FUNCTION_BLOCK "FB_GRAPH_PressDemoAuto"   // FB100, GRAPH
VERSION : 0.1
// stored: AcknowledgeErrorsRequired true, AutoNumber true, GraphVersion 6.0, InitialValuesAcquisition false, IsIECCheckEnabled false, LanguageInNetworks LAD, LockOperatingMode false, PermanentILProcessingInMANMode false, SetENOAutomatically false, SkipSteps false, UDAEnableTagReadback false, WithAlarmHandling true
   // inherited from GRAPH_BASE
   VAR
      OFF_SQ_BASE : Bool;
   END_VAR
   VAR_INPUT
      OFF_SQ { ExternalAccessible := 'False'; ExternalVisible := 'False'; ExternalWritable := 'False'} : Bool := false;   // Turn sequence off
      INIT_SQ { ExternalAccessible := 'False'; ExternalVisible := 'False'; ExternalWritable := 'False'} : Bool := false;   // Set sequence to initial state
      ACK_EF { ExternalAccessible := 'False'; ExternalVisible := 'False'; ExternalWritable := 'False'} : Bool := false;   // Acknowledge all errors and faults
      S_PREV { ExternalAccessible := 'False'; ExternalVisible := 'False'; ExternalWritable := 'False'} : Bool := false;   // Output previous step in parameter S_NO
      S_NEXT { ExternalAccessible := 'False'; ExternalVisible := 'False'; ExternalWritable := 'False'} : Bool := false;   // Indicate next step in parameter S_NO
      SW_AUTO { ExternalAccessible := 'False'; ExternalVisible := 'False'; ExternalWritable := 'False'} : Bool := false;   // Automatic mode
      SW_TAP { ExternalAccessible := 'False'; ExternalVisible := 'False'; ExternalWritable := 'False'} : Bool := false;   // Semiautomatic/switch with transition
      SW_TOP { ExternalAccessible := 'False'; ExternalVisible := 'False'; ExternalWritable := 'False'} : Bool := false;   // Semiautomatic/ignore transition
      SW_MAN { ExternalAccessible := 'False'; ExternalVisible := 'False'; ExternalWritable := 'False'} : Bool := false;   // Manual mode
      S_SEL { ExternalAccessible := 'False'; ExternalVisible := 'False'; ExternalWritable := 'False'} : Int := 0;   // Select step to be output to S_NO
      S_ON { ExternalAccessible := 'False'; ExternalVisible := 'False'; ExternalWritable := 'False'} : Bool := false;   // Activate step indicated in S_NO
      S_OFF { ExternalAccessible := 'False'; ExternalVisible := 'False'; ExternalWritable := 'False'} : Bool := false;   // Disable step indicated in S_NO
      T_PUSH { ExternalAccessible := 'False'; ExternalVisible := 'False'; ExternalWritable := 'False'} : Bool := false;   // Enable transition to switch in semi automatic mode
      Run : Bool;
      Reset : Bool;
      OwnerIndex : DInt;
      Delta : Time;
      TransferSettleTime : Time;
      PartQuality : Bool;
      RequireTwoHandStart : Bool;
      SourcePath : String[80];
      PartPresent : Bool;
      AirPressureOk : Bool;
      TwoHandHeld : Bool;
      StartPulse : Bool;
      PressSettleTime : Time;
   END_VAR
   VAR_OUTPUT
      S_NO { ExternalAccessible := 'False'; ExternalVisible := 'False'; ExternalWritable := 'False'} : Int := 0;   // Step number
      S_MORE { ExternalAccessible := 'False'; ExternalVisible := 'False'; ExternalWritable := 'False'} : Bool := false;   // More steps are available and can be shown in S_NO
      S_ACTIVE { ExternalAccessible := 'False'; ExternalVisible := 'False'; ExternalWritable := 'False'} : Bool := false;   // Step indicated in S_NO is active
      ERR_FLT { ExternalAccessible := 'False'; ExternalVisible := 'False'; ExternalWritable := 'False'} : Bool := false;   // Interlock or supervision group error
      AUTO_ON { ExternalAccessible := 'False'; ExternalVisible := 'False'; ExternalWritable := 'False'} : Bool := false;   // Automatic mode is active
      TAP_ON { ExternalAccessible := 'False'; ExternalVisible := 'False'; ExternalWritable := 'False'} : Bool := false;   // Semiautomatic mode/step with transition enabled
      TOP_ON { ExternalAccessible := 'False'; ExternalVisible := 'False'; ExternalWritable := 'False'} : Bool := false;   // Semiautomatic mode/ignore transition enabled
      MAN_ON { ExternalAccessible := 'False'; ExternalVisible := 'False'; ExternalWritable := 'False'} : Bool := false;   // Manual mode is active
   END_VAR
   VAR_IN_OUT
      PressRam : "FB_CylinderCM";
      Door : "FB_CylinderCM";
      PartSlide : "FB_CylinderCM";
      HostCore : "FRK_Core";
      HostUnit : "FRK_Unit";
      HostStatus : "ST_ModuleStatus";
      HostPart : "ST_PartContext";
      HostAlarmLog : "FRK_AlarmLog";
      Seq : "FRK_SequenceCtx";
      Row1 : "FRK_SequenceRow";
      Row2 : "FRK_SequenceRow";
      Row3 : "FRK_SequenceRow";
      Row4 : "FRK_SequenceRow";
      Row5 : "FRK_SequenceRow";
      Row6 : "FRK_SequenceRow";
      Row7 : "FRK_SequenceRow";
      Row8 : "FRK_SequenceRow";
      Row9 : "FRK_SequenceRow";
      Row10 : "FRK_SequenceRow";
      Row11 : "FRK_SequenceRow";
      Row12 : "FRK_SequenceRow";
      Row13 : "FRK_SequenceRow";
      Row14 : "FRK_SequenceRow";
      Row15 : "FRK_SequenceRow";
      Row16 : "FRK_SequenceRow";
      Ready1 { ExternalAccessible := 'False'; ExternalVisible := 'False'; ExternalWritable := 'False'} : Bool;
      Ready2 { ExternalAccessible := 'False'; ExternalVisible := 'False'; ExternalWritable := 'False'} : Bool;
      Ready3 { ExternalAccessible := 'False'; ExternalVisible := 'False'; ExternalWritable := 'False'} : Bool;
      Ready4 { ExternalAccessible := 'False'; ExternalVisible := 'False'; ExternalWritable := 'False'} : Bool;
      Ready5 { ExternalAccessible := 'False'; ExternalVisible := 'False'; ExternalWritable := 'False'} : Bool;
      Cycle : "ST_PressDemoCycle";
      LoadDone { ExternalAccessible := 'False'; ExternalVisible := 'False'; ExternalWritable := 'False'} : Bool;
      Branch1 : "FRK_SequenceCtx";
      Branch2 : "FRK_SequenceCtx";
      Row17 : "FRK_SequenceRow";
      Row18 : "FRK_SequenceRow";
      Row19 : "FRK_SequenceRow";
   END_VAR
BEGIN
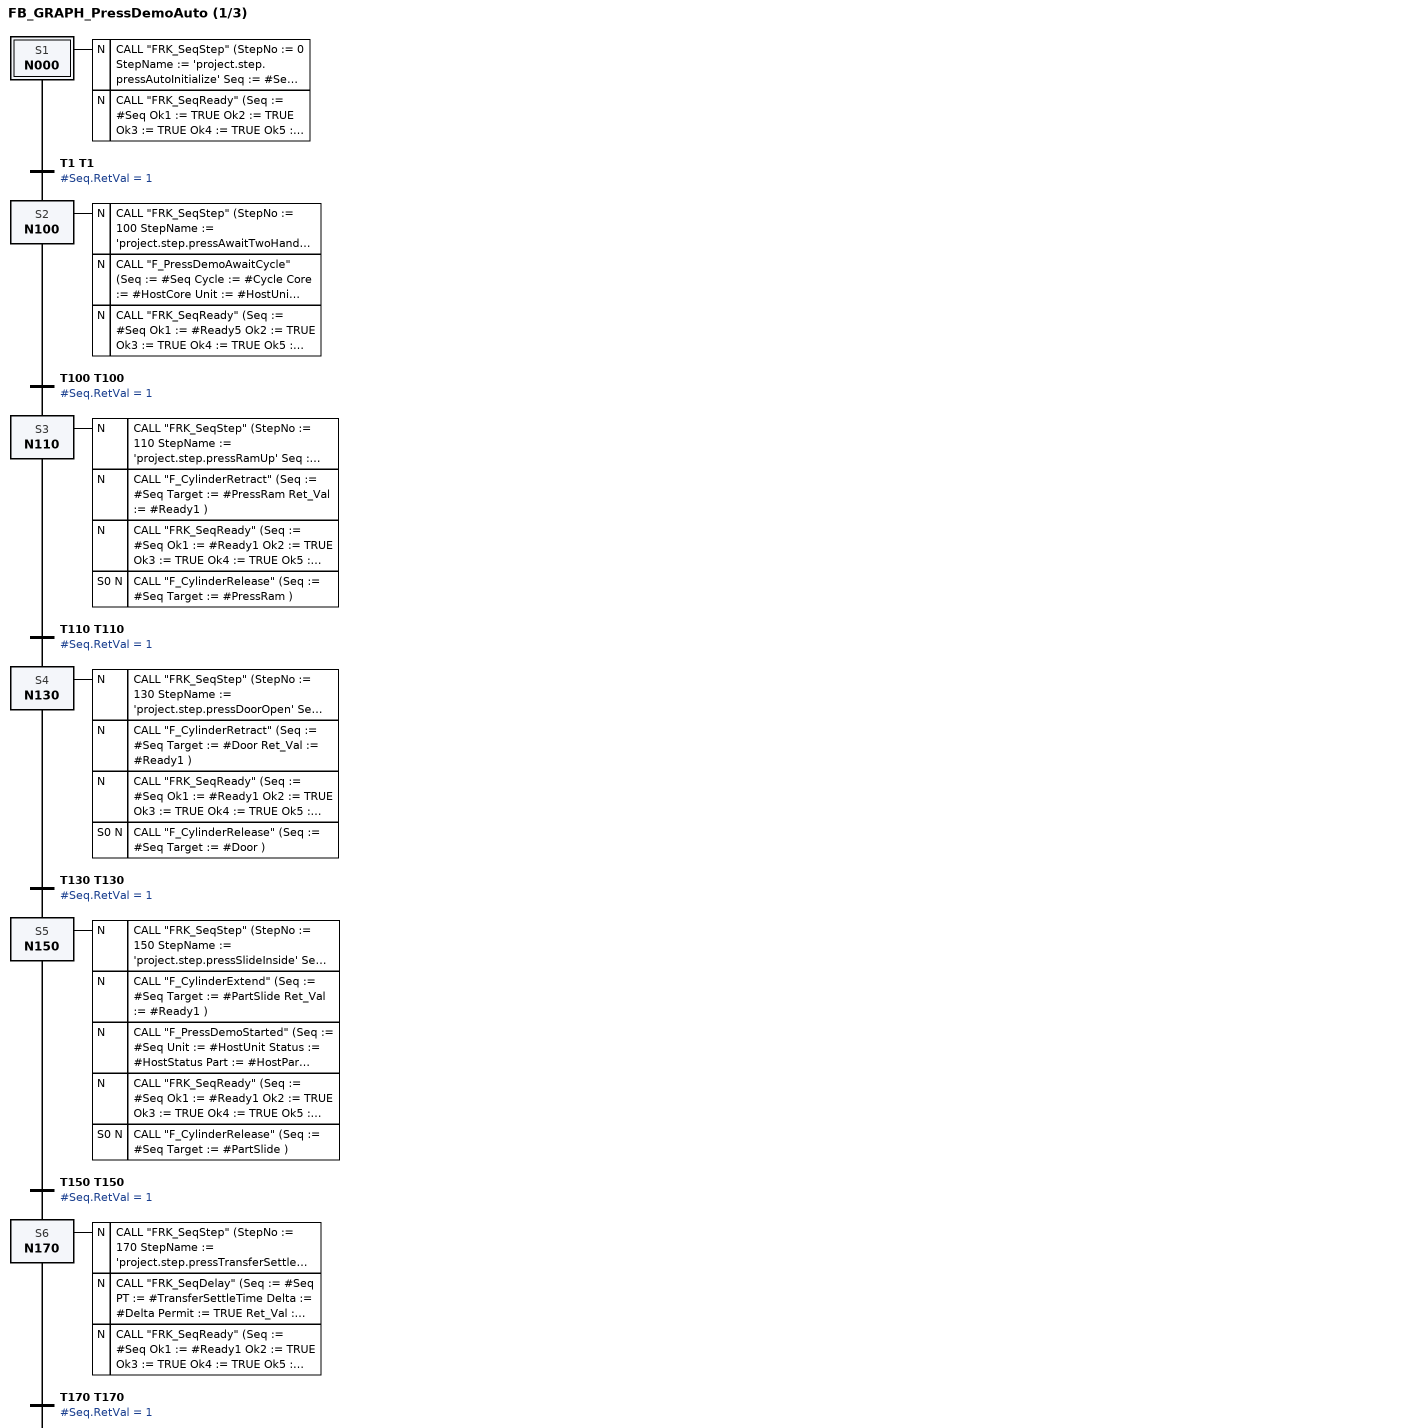
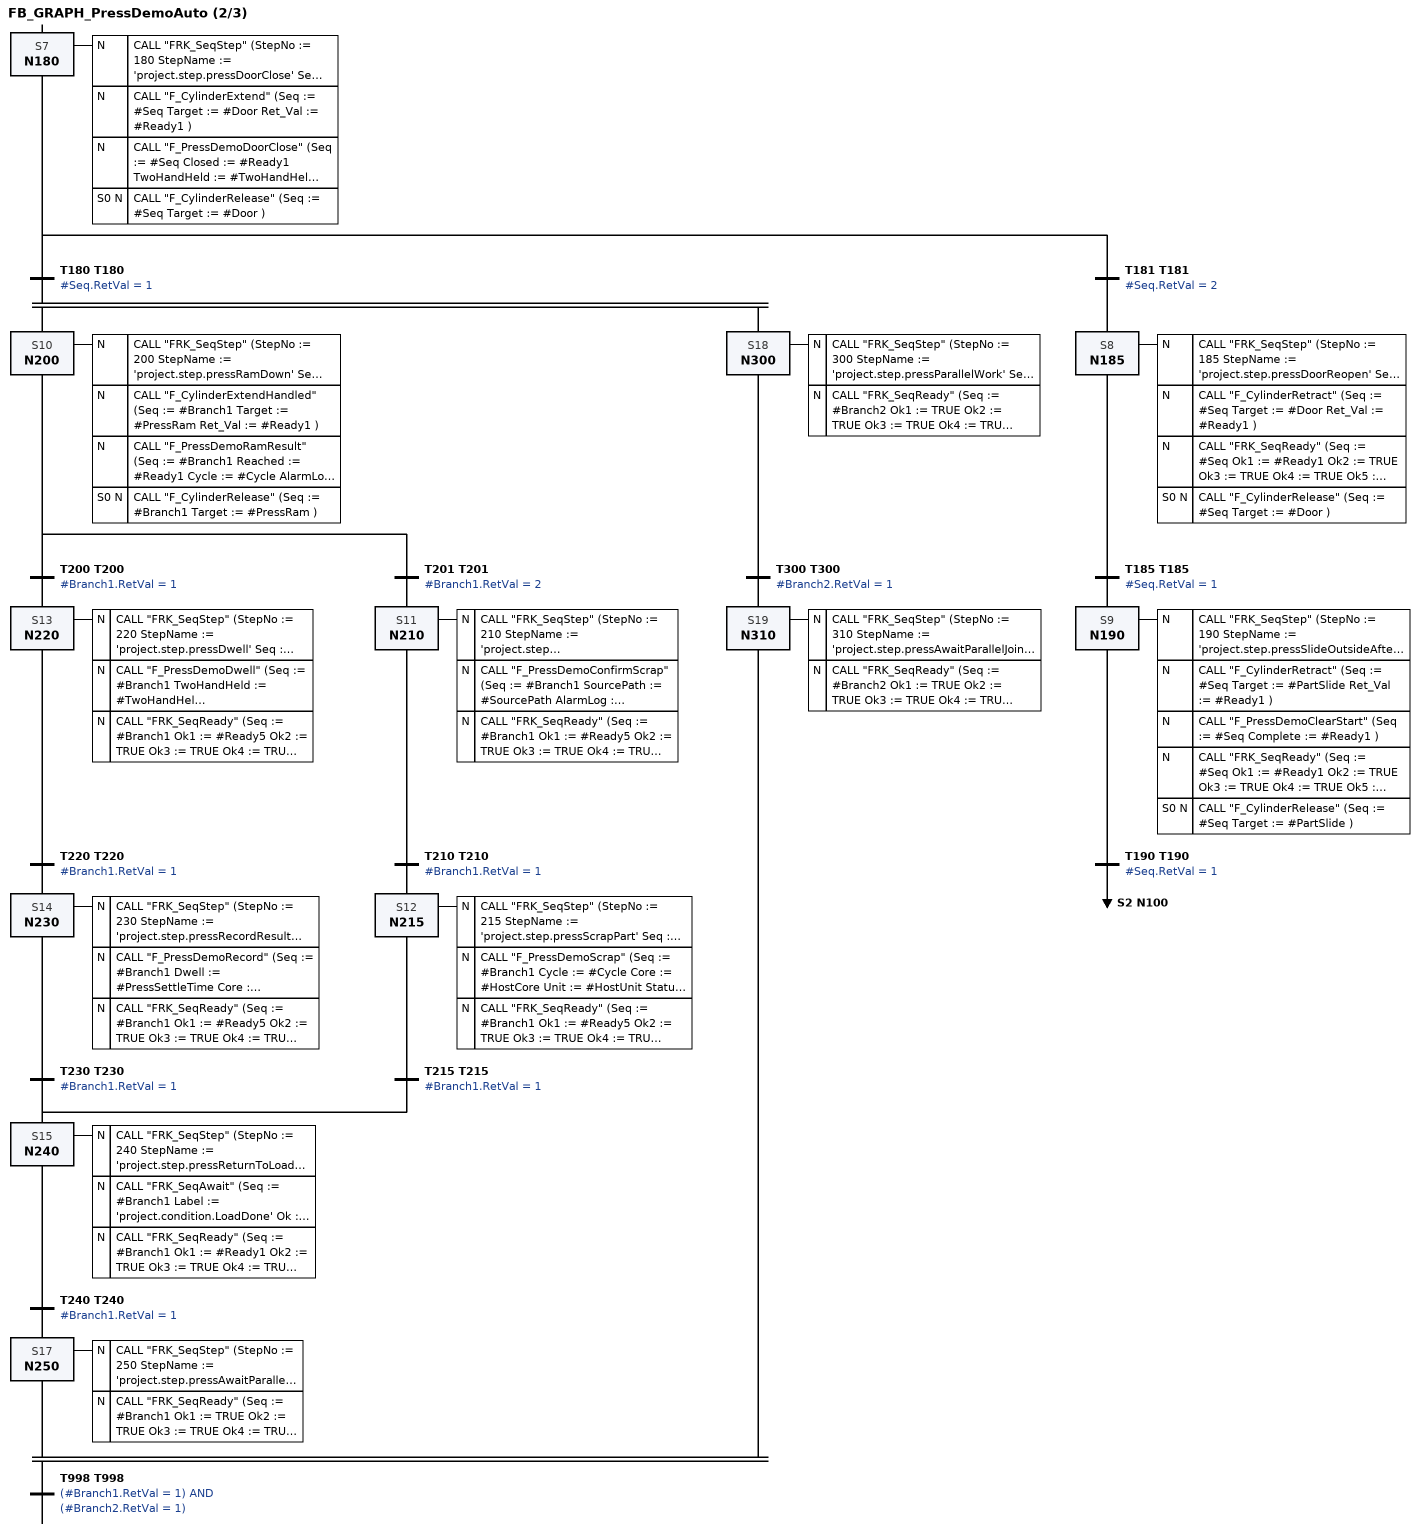
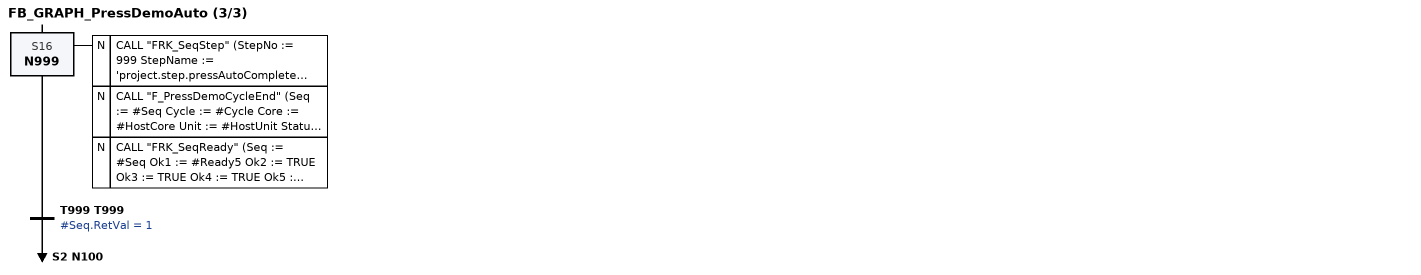
   // sequencer 1
   INITIAL_STEP N000:   // S1, max time T#10S, warning time T#7S
              N    CALL "FRK_SeqStep" 
                   (StepNo := 0
                   StepName := 'project.step.pressAutoInitialize'
                   Seq := #Seq
                   Row := #Row1
                   )
              N    CALL "FRK_SeqReady" 
                   (Seq := #Seq
                   Ok1 := TRUE
                   Ok2 := TRUE
                   Ok3 := TRUE
                   Ok4 := TRUE
                   Ok5 := TRUE
                   )
   END_STEP
   TRANSITION T1 FROM N000 TO N100   // T1
      := #Seq.RetVal = 1;
   END_TRANSITION
   STEP N100:   // S2, max time T#10S, warning time T#7S
              N    CALL "FRK_SeqStep" 
                   (StepNo := 100
                   StepName := 'project.step.pressAwaitTwoHand'
                   Seq := #Seq
                   Row := #Row2
                   )
              N    CALL "F_PressDemoAwaitCycle" 
                   (Seq := #Seq
                   Cycle := #Cycle
                   Core := #HostCore
                   Unit := #HostUnit
                   Status := #HostStatus
                   Part := #HostPart
                   AlarmLog := #HostAlarmLog
                   PartPresent := #PartPresent
                   PartQuality := #PartQuality
                   AirPressureOk := #AirPressureOk
                   RequireTwoHandStart := #RequireTwoHandStart
                   Ret_Val := #Ready5
                   )
              N    CALL "FRK_SeqReady" 
                   (Seq := #Seq
                   Ok1 := #Ready5
                   Ok2 := TRUE
                   Ok3 := TRUE
                   Ok4 := TRUE
                   Ok5 := TRUE
                   )
   END_STEP
   TRANSITION T100 FROM N100 TO N110   // T100
      := #Seq.RetVal = 1;
   END_TRANSITION
   STEP N110:   // S3, max time T#10S, warning time T#7S
              N    CALL "FRK_SeqStep" 
                   (StepNo := 110
                   StepName := 'project.step.pressRamUp'
                   Seq := #Seq
                   Row := #Row3
                   )
              N    CALL "F_CylinderRetract" 
                   (Seq := #Seq
                   Target := #PressRam
                   Ret_Val := #Ready1
                   )
              N    CALL "FRK_SeqReady" 
                   (Seq := #Seq
                   Ok1 := #Ready1
                   Ok2 := TRUE
                   Ok3 := TRUE
                   Ok4 := TRUE
                   Ok5 := TRUE
                   )
          S0  N    CALL "F_CylinderRelease" 
                   (Seq := #Seq
                   Target := #PressRam
                   )
   END_STEP
   TRANSITION T110 FROM N110 TO N130   // T110
      := #Seq.RetVal = 1;
   END_TRANSITION
   STEP N130:   // S4, max time T#10S, warning time T#7S
              N    CALL "FRK_SeqStep" 
                   (StepNo := 130
                   StepName := 'project.step.pressDoorOpen'
                   Seq := #Seq
                   Row := #Row4
                   )
              N    CALL "F_CylinderRetract" 
                   (Seq := #Seq
                   Target := #Door
                   Ret_Val := #Ready1
                   )
              N    CALL "FRK_SeqReady" 
                   (Seq := #Seq
                   Ok1 := #Ready1
                   Ok2 := TRUE
                   Ok3 := TRUE
                   Ok4 := TRUE
                   Ok5 := TRUE
                   )
          S0  N    CALL "F_CylinderRelease" 
                   (Seq := #Seq
                   Target := #Door
                   )
   END_STEP
   TRANSITION T130 FROM N130 TO N150   // T130
      := #Seq.RetVal = 1;
   END_TRANSITION
   STEP N150:   // S5, max time T#10S, warning time T#7S
              N    CALL "FRK_SeqStep" 
                   (StepNo := 150
                   StepName := 'project.step.pressSlideInside'
                   Seq := #Seq
                   Row := #Row5
                   )
              N    CALL "F_CylinderExtend" 
                   (Seq := #Seq
                   Target := #PartSlide
                   Ret_Val := #Ready1
                   )
              N    CALL "F_PressDemoStarted" 
                   (Seq := #Seq
                   Unit := #HostUnit
                   Status := #HostStatus
                   Part := #HostPart
                   AlarmLog := #HostAlarmLog
                   )
              N    CALL "FRK_SeqReady" 
                   (Seq := #Seq
                   Ok1 := #Ready1
                   Ok2 := TRUE
                   Ok3 := TRUE
                   Ok4 := TRUE
                   Ok5 := TRUE
                   )
          S0  N    CALL "F_CylinderRelease" 
                   (Seq := #Seq
                   Target := #PartSlide
                   )
   END_STEP
   TRANSITION T150 FROM N150 TO N170   // T150
      := #Seq.RetVal = 1;
   END_TRANSITION
   STEP N170:   // S6, max time T#10S, warning time T#7S
              N    CALL "FRK_SeqStep" 
                   (StepNo := 170
                   StepName := 'project.step.pressTransferSettle'
                   Seq := #Seq
                   Row := #Row6
                   )
              N    CALL "FRK_SeqDelay" 
                   (Seq := #Seq
                   PT := #TransferSettleTime
                   Delta := #Delta
                   Permit := TRUE
                   Ret_Val := #Ready1
                   )
              N    CALL "FRK_SeqReady" 
                   (Seq := #Seq
                   Ok1 := #Ready1
                   Ok2 := TRUE
                   Ok3 := TRUE
                   Ok4 := TRUE
                   Ok5 := TRUE
                   )
   END_STEP
   TRANSITION T170 FROM N170 TO N180   // T170
      := #Seq.RetVal = 1;
   END_TRANSITION
   STEP N180:   // S7, max time T#10S, warning time T#7S
              N    CALL "FRK_SeqStep" 
                   (StepNo := 180
                   StepName := 'project.step.pressDoorClose'
                   Seq := #Seq
                   Row := #Row7
                   )
              N    CALL "F_CylinderExtend" 
                   (Seq := #Seq
                   Target := #Door
                   Ret_Val := #Ready1
                   )
              N    CALL "F_PressDemoDoorClose" 
                   (Seq := #Seq
                   Closed := #Ready1
                   TwoHandHeld := #TwoHandHeld
                   RequireTwoHandStart := #RequireTwoHandStart
                   SourcePath := #SourcePath
                   AlarmLog := #HostAlarmLog
                   )
          S0  N    CALL "F_CylinderRelease" 
                   (Seq := #Seq
                   Target := #Door
                   )
   END_STEP
   TRANSITION T180 FROM N180 TO (N200, N300)   // T180
      := #Seq.RetVal = 1;
   END_TRANSITION
   TRANSITION T181 FROM N180 TO N185   // T181
      := #Seq.RetVal = 2;
   END_TRANSITION
   STEP N185:   // S8, max time T#10S, warning time T#7S
              N    CALL "FRK_SeqStep" 
                   (StepNo := 185
                   StepName := 'project.step.pressDoorReopen'
                   Seq := #Seq
                   Row := #Row8
                   )
              N    CALL "F_CylinderRetract" 
                   (Seq := #Seq
                   Target := #Door
                   Ret_Val := #Ready1
                   )
              N    CALL "FRK_SeqReady" 
                   (Seq := #Seq
                   Ok1 := #Ready1
                   Ok2 := TRUE
                   Ok3 := TRUE
                   Ok4 := TRUE
                   Ok5 := TRUE
                   )
          S0  N    CALL "F_CylinderRelease" 
                   (Seq := #Seq
                   Target := #Door
                   )
   END_STEP
   TRANSITION T185 FROM N185 TO N190   // T185
      := #Seq.RetVal = 1;
   END_TRANSITION
   STEP N190:   // S9, max time T#10S, warning time T#7S
              N    CALL "FRK_SeqStep" 
                   (StepNo := 190
                   StepName := 'project.step.pressSlideOutsideAfterAbort'
                   Seq := #Seq
                   Row := #Row9
                   )
              N    CALL "F_CylinderRetract" 
                   (Seq := #Seq
                   Target := #PartSlide
                   Ret_Val := #Ready1
                   )
              N    CALL "F_PressDemoClearStart" 
                   (Seq := #Seq
                   Complete := #Ready1
                   )
              N    CALL "FRK_SeqReady" 
                   (Seq := #Seq
                   Ok1 := #Ready1
                   Ok2 := TRUE
                   Ok3 := TRUE
                   Ok4 := TRUE
                   Ok5 := TRUE
                   )
          S0  N    CALL "F_CylinderRelease" 
                   (Seq := #Seq
                   Target := #PartSlide
                   )
   END_STEP
   TRANSITION T190 FROM N190 TO N100   // T190, jump
      := #Seq.RetVal = 1;
   END_TRANSITION
   STEP N200:   // S10, max time T#10S, warning time T#7S
              N    CALL "FRK_SeqStep" 
                   (StepNo := 200
                   StepName := 'project.step.pressRamDown'
                   Seq := #Branch1
                   Row := #Row10
                   )
              N    CALL "F_CylinderExtendHandled" 
                   (Seq := #Branch1
                   Target := #PressRam
                   Ret_Val := #Ready1
                   )
              N    CALL "F_PressDemoRamResult" 
                   (Seq := #Branch1
                   Reached := #Ready1
                   Cycle := #Cycle
                   AlarmLog := #HostAlarmLog
                   )
          S0  N    CALL "F_CylinderRelease" 
                   (Seq := #Branch1
                   Target := #PressRam
                   )
   END_STEP
   TRANSITION T200 FROM N200 TO N220   // T200
      := #Branch1.RetVal = 1;
   END_TRANSITION
   TRANSITION T201 FROM N200 TO N210   // T201
      := #Branch1.RetVal = 2;
   END_TRANSITION
   STEP N210:   // S11, max time T#10S, warning time T#7S
              N    CALL "FRK_SeqStep" 
                   (StepNo := 210
                   StepName := 'project.step.pressNotReachedConfirm'
                   Seq := #Branch1
                   Row := #Row11
                   )
              N    CALL "F_PressDemoConfirmScrap" 
                   (Seq := #Branch1
                   SourcePath := #SourcePath
                   AlarmLog := #HostAlarmLog
                   Ret_Val := #Ready5
                   )
              N    CALL "FRK_SeqReady" 
                   (Seq := #Branch1
                   Ok1 := #Ready5
                   Ok2 := TRUE
                   Ok3 := TRUE
                   Ok4 := TRUE
                   Ok5 := TRUE
                   )
   END_STEP
   TRANSITION T210 FROM N210 TO N215   // T210
      := #Branch1.RetVal = 1;
   END_TRANSITION
   STEP N215:   // S12, max time T#10S, warning time T#7S
              N    CALL "FRK_SeqStep" 
                   (StepNo := 215
                   StepName := 'project.step.pressScrapPart'
                   Seq := #Branch1
                   Row := #Row12
                   )
              N    CALL "F_PressDemoScrap" 
                   (Seq := #Branch1
                   Cycle := #Cycle
                   Core := #HostCore
                   Unit := #HostUnit
                   Status := #HostStatus
                   Part := #HostPart
                   AlarmLog := #HostAlarmLog
                   Ret_Val := #Ready5
                   )
              N    CALL "FRK_SeqReady" 
                   (Seq := #Branch1
                   Ok1 := #Ready5
                   Ok2 := TRUE
                   Ok3 := TRUE
                   Ok4 := TRUE
                   Ok5 := TRUE
                   )
   END_STEP
   TRANSITION T215 FROM N215 TO N240   // T215
      := #Branch1.RetVal = 1;
   END_TRANSITION
   STEP N220:   // S13, max time T#10S, warning time T#7S
              N    CALL "FRK_SeqStep" 
                   (StepNo := 220
                   StepName := 'project.step.pressDwell'
                   Seq := #Branch1
                   Row := #Row13
                   )
              N    CALL "F_PressDemoDwell" 
                   (Seq := #Branch1
                   TwoHandHeld := #TwoHandHeld
                   RequireTwoHandStart := #RequireTwoHandStart
                   PT := #PressSettleTime
                   Delta := #Delta
                   PressRam := #PressRam
                   Ret_Val := #Ready5
                   )
              N    CALL "FRK_SeqReady" 
                   (Seq := #Branch1
                   Ok1 := #Ready5
                   Ok2 := TRUE
                   Ok3 := TRUE
                   Ok4 := TRUE
                   Ok5 := TRUE
                   )
   END_STEP
   TRANSITION T220 FROM N220 TO N230   // T220
      := #Branch1.RetVal = 1;
   END_TRANSITION
   STEP N230:   // S14, max time T#10S, warning time T#7S
              N    CALL "FRK_SeqStep" 
                   (StepNo := 230
                   StepName := 'project.step.pressRecordResult'
                   Seq := #Branch1
                   Row := #Row14
                   )
              N    CALL "F_PressDemoRecord" 
                   (Seq := #Branch1
                   Dwell := #PressSettleTime
                   Core := #HostCore
                   Status := #HostStatus
                   Part := #HostPart
                   Ret_Val := #Ready5
                   )
              N    CALL "FRK_SeqReady" 
                   (Seq := #Branch1
                   Ok1 := #Ready5
                   Ok2 := TRUE
                   Ok3 := TRUE
                   Ok4 := TRUE
                   Ok5 := TRUE
                   )
   END_STEP
   TRANSITION T230 FROM N230 TO N240   // T230
      := #Branch1.RetVal = 1;
   END_TRANSITION
   STEP N240:   // S15, max time T#10S, warning time T#7S
              N    CALL "FRK_SeqStep" 
                   (StepNo := 240
                   StepName := 'project.step.pressReturnToLoad'
                   Seq := #Branch1
                   Row := #Row15
                   )
              N    CALL "FRK_SeqAwait" 
                   (Seq := #Branch1
                   Label := 'project.condition.LoadDone'
                   Ok := #LoadDone
                   Ret_Val := #Ready1
                   )
              N    CALL "FRK_SeqReady" 
                   (Seq := #Branch1
                   Ok1 := #Ready1
                   Ok2 := TRUE
                   Ok3 := TRUE
                   Ok4 := TRUE
                   Ok5 := TRUE
                   )
   END_STEP
   TRANSITION T240 FROM N240 TO N250   // T240
      := #Branch1.RetVal = 1;
   END_TRANSITION
   STEP N999:   // S16, max time T#10S, warning time T#7S
              N    CALL "FRK_SeqStep" 
                   (StepNo := 999
                   StepName := 'project.step.pressAutoComplete'
                   Seq := #Seq
                   Row := #Row16
                   )
              N    CALL "F_PressDemoCycleEnd" 
                   (Seq := #Seq
                   Cycle := #Cycle
                   Core := #HostCore
                   Unit := #HostUnit
                   Status := #HostStatus
                   Part := #HostPart
                   AlarmLog := #HostAlarmLog
                   Ret_Val := #Ready5
                   )
              N    CALL "FRK_SeqReady" 
                   (Seq := #Seq
                   Ok1 := #Ready5
                   Ok2 := TRUE
                   Ok3 := TRUE
                   Ok4 := TRUE
                   Ok5 := TRUE
                   )
   END_STEP
   TRANSITION T999 FROM N999 TO N100   // T999, jump
      := #Seq.RetVal = 1;
   END_TRANSITION
   STEP N250:   // S17, max time T#10S, warning time T#7S
              N    CALL "FRK_SeqStep" 
                   (StepNo := 250
                   StepName := 'project.step.pressAwaitParallelBranch'
                   Seq := #Branch1
                   Row := #Row17
                   )
              N    CALL "FRK_SeqReady" 
                   (Seq := #Branch1
                   Ok1 := TRUE
                   Ok2 := TRUE
                   Ok3 := TRUE
                   Ok4 := TRUE
                   Ok5 := TRUE
                   )
   END_STEP
   STEP N300:   // S18, max time T#10S, warning time T#7S
              N    CALL "FRK_SeqStep" 
                   (StepNo := 300
                   StepName := 'project.step.pressParallelWork'
                   Seq := #Branch2
                   Row := #Row18
                   )
              N    CALL "FRK_SeqReady" 
                   (Seq := #Branch2
                   Ok1 := TRUE
                   Ok2 := TRUE
                   Ok3 := TRUE
                   Ok4 := TRUE
                   Ok5 := TRUE
                   )
   END_STEP
   TRANSITION T300 FROM N300 TO N310   // T300
      := #Branch2.RetVal = 1;
   END_TRANSITION
   STEP N310:   // S19, max time T#10S, warning time T#7S
              N    CALL "FRK_SeqStep" 
                   (StepNo := 310
                   StepName := 'project.step.pressAwaitParallelJoin'
                   Seq := #Branch2
                   Row := #Row19
                   )
              N    CALL "FRK_SeqReady" 
                   (Seq := #Branch2
                   Ok1 := TRUE
                   Ok2 := TRUE
                   Ok3 := TRUE
                   Ok4 := TRUE
                   Ok5 := TRUE
                   )
   END_STEP
   TRANSITION T998 FROM (N250, N310) TO N999   // T998
      := (#Branch1.RetVal = 1) AND (#Branch2.RetVal = 1);
   END_TRANSITION
END_FUNCTION_BLOCK

FUNCTION_BLOCK "FB_PressDemoLoadPosition"   // FB2, SCL
{ S7_Optimized_Access := 'TRUE' }
VERSION : 0.1
// stored: AutoNumber true, IsIECCheckEnabled false, IsRetainMemResEnabled false, MemoryReserve 100, SetENOAutomatically false, UDAEnableTagReadback false
   VAR_INPUT
      Run : Bool;
      Reset : Bool;
      OwnerIndex : DInt;
      Delta : Time;
   END_VAR
   VAR_IN_OUT
      PressRam : "FB_CylinderCM";
      Door : "FB_CylinderCM";
      PartSlide : "FB_CylinderCM";
   END_VAR
   VAR
      Seq { ExternalWritable := 'False'; S7_SetPoint := 'True'} : "FRK_SequenceCtx";
      Row1 { ExternalWritable := 'False'; S7_SetPoint := 'True'} : "FRK_SequenceRow";
      Row2 { ExternalWritable := 'False'; S7_SetPoint := 'True'} : "FRK_SequenceRow";
      Row3 { ExternalWritable := 'False'; S7_SetPoint := 'True'} : "FRK_SequenceRow";
      Row4 { ExternalWritable := 'False'; S7_SetPoint := 'True'} : "FRK_SequenceRow";
      At240 { ExternalAccessible := 'False'; ExternalVisible := 'False'; ExternalWritable := 'False'} : Bool;
      At260 { ExternalAccessible := 'False'; ExternalVisible := 'False'; ExternalWritable := 'False'} : Bool;
      At280 { ExternalAccessible := 'False'; ExternalVisible := 'False'; ExternalWritable := 'False'} : Bool;
      At300 { ExternalAccessible := 'False'; ExternalVisible := 'False'; ExternalWritable := 'False'} : Bool;
      Ready1 { ExternalAccessible := 'False'; ExternalVisible := 'False'; ExternalWritable := 'False'} : Bool;
      Ready2 { ExternalAccessible := 'False'; ExternalVisible := 'False'; ExternalWritable := 'False'} : Bool;
      Ready3 { ExternalAccessible := 'False'; ExternalVisible := 'False'; ExternalWritable := 'False'} : Bool;
      Ready4 { ExternalAccessible := 'False'; ExternalVisible := 'False'; ExternalWritable := 'False'} : Bool;
      Ready5 { ExternalAccessible := 'False'; ExternalVisible := 'False'; ExternalWritable := 'False'} : Bool;
      Advance { ExternalAccessible := 'False'; ExternalVisible := 'False'; ExternalWritable := 'False'} : Bool;
   END_VAR
BEGIN

   "FRK_SeqBegin"(Run := #Run,
                  Reset := #Reset,
                  OwnerIndex := #OwnerIndex,
                  ChainIndex := 3,
                  BranchIndex := 1,
                  Delta := #Delta,
                  Seq := #Seq);
   "FRK_SeqInitial"(Seq := #Seq,
                    InitialStep := 240);
   "F_CylinderSequenceLease"(Seq := #Seq,
                             Target := #PressRam);
   "F_CylinderSequenceLease"(Seq := #Seq,
                             Target := #Door);
   "F_CylinderSequenceLease"(Seq := #Seq,
                             Target := #PartSlide);
   CASE #Seq.ScanStep OF
       240:
           IF #Seq.Running AND NOT #Seq.Error THEN
               "FRK_SeqStep"(StepNo := 240,
                             StepName := 'project.step.pressReturnRam',
                             Seq := #Seq,
                             Row := #Row1);
               #Ready1 := "F_CylinderRetract"(Seq := #Seq, Target := #PressRam);
               "FRK_SeqReady"(Seq := #Seq,
                              Ok1 := #Ready1,
                              Ok2 := TRUE,
                              Ok3 := TRUE,
                              Ok4 := TRUE,
                              Ok5 := TRUE);
               "FRK_SeqRoute"(Seq := #Seq,
                              OnAdvance := 260,
                              OnJump1 := -1);
           END_IF;
       260:
           IF #Seq.Running AND NOT #Seq.Error THEN
               "FRK_SeqStep"(StepNo := 260,
                             StepName := 'project.step.pressReturnDoor',
                             Seq := #Seq,
                             Row := #Row2);
               #Ready1 := "F_CylinderRetract"(Seq := #Seq, Target := #Door);
               "FRK_SeqReady"(Seq := #Seq,
                              Ok1 := #Ready1,
                              Ok2 := TRUE,
                              Ok3 := TRUE,
                              Ok4 := TRUE,
                              Ok5 := TRUE);
               "FRK_SeqRoute"(Seq := #Seq,
                              OnAdvance := 280,
                              OnJump1 := -1);
           END_IF;
       280:
           IF #Seq.Running AND NOT #Seq.Error THEN
               "FRK_SeqStep"(StepNo := 280,
                             StepName := 'project.step.pressReturnSlide',
                             Seq := #Seq,
                             Row := #Row3);
               #Ready1 := "F_CylinderRetract"(Seq := #Seq, Target := #PartSlide);
               "FRK_SeqReady"(Seq := #Seq,
                              Ok1 := #Ready1,
                              Ok2 := TRUE,
                              Ok3 := TRUE,
                              Ok4 := TRUE,
                              Ok5 := TRUE);
               "FRK_SeqRoute"(Seq := #Seq,
                              OnAdvance := 300,
                              OnJump1 := -1);
           END_IF;
       300:
           IF #Seq.Running AND NOT #Seq.Error THEN
               "FRK_SeqStep"(StepNo := 300,
                             StepName := 'project.step.pressLoadPositionComplete',
                             Seq := #Seq,
                             Row := #Row4);
               "FRK_SeqComplete"(Seq := #Seq);
           END_IF;
       ELSE
           #Seq.Error := TRUE;
           #Seq.ErrorDiagnostic.ReasonCode := 10001;
           #Seq.ErrorDiagnostic.Description := WSTRING#'project.sequence.invalidStep';
   END_CASE;
   "F_CylinderSequenceLease"(Seq := #Seq,
                             Target := #PressRam);
   "F_CylinderSequenceLease"(Seq := #Seq,
                             Target := #Door);
   "F_CylinderSequenceLease"(Seq := #Seq,
                             Target := #PartSlide);
END_FUNCTION_BLOCK

FUNCTION_BLOCK "FB_PressDemoHomeGraphOwner"   // FB11, SCL
{ S7_Optimized_Access := 'TRUE' }
VERSION : 0.1
// stored: AutoNumber true, IsIECCheckEnabled false, IsRetainMemResEnabled false, MemoryReserve 100, SetENOAutomatically false, UDAEnableTagReadback false
   VAR_INPUT
      Run : Bool;
      Reset : Bool;
      OwnerIndex : DInt;
      Delta : Time;
   END_VAR
   VAR_IN_OUT
      PressRam : "FB_CylinderCM";
      Door : "FB_CylinderCM";
      PartSlide : "FB_CylinderCM";
      Chart : "FB_GRAPH_PressDemoHome";
   END_VAR
   VAR
      Seq { ExternalWritable := 'False'; S7_SetPoint := 'True'} : "FRK_SequenceCtx";
      Row1 { ExternalWritable := 'False'; S7_SetPoint := 'True'} : "FRK_SequenceRow";
      Row2 { ExternalWritable := 'False'; S7_SetPoint := 'True'} : "FRK_SequenceRow";
      Row3 { ExternalWritable := 'False'; S7_SetPoint := 'True'} : "FRK_SequenceRow";
      Row4 { ExternalWritable := 'False'; S7_SetPoint := 'True'} : "FRK_SequenceRow";
      At0 { ExternalAccessible := 'False'; ExternalVisible := 'False'; ExternalWritable := 'False'} : Bool;
      At900 { ExternalAccessible := 'False'; ExternalVisible := 'False'; ExternalWritable := 'False'} : Bool;
      At910 { ExternalAccessible := 'False'; ExternalVisible := 'False'; ExternalWritable := 'False'} : Bool;
      At999 { ExternalAccessible := 'False'; ExternalVisible := 'False'; ExternalWritable := 'False'} : Bool;
      Ready1 { ExternalAccessible := 'False'; ExternalVisible := 'False'; ExternalWritable := 'False'} : Bool;
      Ready2 { ExternalAccessible := 'False'; ExternalVisible := 'False'; ExternalWritable := 'False'} : Bool;
      Ready3 { ExternalAccessible := 'False'; ExternalVisible := 'False'; ExternalWritable := 'False'} : Bool;
      Ready4 { ExternalAccessible := 'False'; ExternalVisible := 'False'; ExternalWritable := 'False'} : Bool;
      Ready5 { ExternalAccessible := 'False'; ExternalVisible := 'False'; ExternalWritable := 'False'} : Bool;
      Advance { ExternalAccessible := 'False'; ExternalVisible := 'False'; ExternalWritable := 'False'} : Bool;
   END_VAR
BEGIN

   "FRK_SeqBegin"(Run := #Run,
                  Reset := #Reset,
                  OwnerIndex := #OwnerIndex,
                  ChainIndex := 2,
                  BranchIndex := 0,
                  Delta := #Delta,
                  Seq := #Seq);
   "F_CylinderSequenceLease"(Seq := #Seq,
                             Target := #PressRam);
   "F_CylinderSequenceLease"(Seq := #Seq,
                             Target := #Door);
   "F_CylinderSequenceLease"(Seq := #Seq,
                             Target := #PartSlide);
   #Chart(Run := #Run,
          Reset := #Reset,
          OwnerIndex := #OwnerIndex,
          Delta := #Delta,
          PressRam := #PressRam,
          Door := #Door,
          PartSlide := #PartSlide,
          Seq := #Seq,
          Row1 := #Row1,
          Row2 := #Row2,
          Row3 := #Row3,
          Row4 := #Row4,
          Ready1 := #Ready1,
          Ready2 := #Ready2,
          Ready3 := #Ready3,
          Ready4 := #Ready4,
          Ready5 := #Ready5,
          INIT_SQ := #Seq.Restart,
          OFF_SQ := NOT #Seq.Running);
   "F_CylinderSequenceLease"(Seq := #Seq,
                             Target := #PressRam);
   "F_CylinderSequenceLease"(Seq := #Seq,
                             Target := #Door);
   "F_CylinderSequenceLease"(Seq := #Seq,
                             Target := #PartSlide);
END_FUNCTION_BLOCK

FUNCTION_BLOCK "FB_GRAPH_PressDemoHome"   // FB101, GRAPH
VERSION : 0.1
// stored: AcknowledgeErrorsRequired true, AutoNumber true, GraphVersion 6.0, InitialValuesAcquisition false, IsIECCheckEnabled false, LanguageInNetworks LAD, LockOperatingMode false, PermanentILProcessingInMANMode false, SetENOAutomatically false, SkipSteps false, UDAEnableTagReadback false, WithAlarmHandling true
   // inherited from GRAPH_BASE
   VAR
      OFF_SQ_BASE : Bool;
   END_VAR
   VAR_INPUT
      OFF_SQ { ExternalAccessible := 'False'; ExternalVisible := 'False'; ExternalWritable := 'False'} : Bool := false;   // Turn sequence off
      INIT_SQ { ExternalAccessible := 'False'; ExternalVisible := 'False'; ExternalWritable := 'False'} : Bool := false;   // Set sequence to initial state
      ACK_EF { ExternalAccessible := 'False'; ExternalVisible := 'False'; ExternalWritable := 'False'} : Bool := false;   // Acknowledge all errors and faults
      S_PREV { ExternalAccessible := 'False'; ExternalVisible := 'False'; ExternalWritable := 'False'} : Bool := false;   // Output previous step in parameter S_NO
      S_NEXT { ExternalAccessible := 'False'; ExternalVisible := 'False'; ExternalWritable := 'False'} : Bool := false;   // Indicate next step in parameter S_NO
      SW_AUTO { ExternalAccessible := 'False'; ExternalVisible := 'False'; ExternalWritable := 'False'} : Bool := false;   // Automatic mode
      SW_TAP { ExternalAccessible := 'False'; ExternalVisible := 'False'; ExternalWritable := 'False'} : Bool := false;   // Semiautomatic/switch with transition
      SW_TOP { ExternalAccessible := 'False'; ExternalVisible := 'False'; ExternalWritable := 'False'} : Bool := false;   // Semiautomatic/ignore transition
      SW_MAN { ExternalAccessible := 'False'; ExternalVisible := 'False'; ExternalWritable := 'False'} : Bool := false;   // Manual mode
      S_SEL { ExternalAccessible := 'False'; ExternalVisible := 'False'; ExternalWritable := 'False'} : Int := 0;   // Select step to be output to S_NO
      S_ON { ExternalAccessible := 'False'; ExternalVisible := 'False'; ExternalWritable := 'False'} : Bool := false;   // Activate step indicated in S_NO
      S_OFF { ExternalAccessible := 'False'; ExternalVisible := 'False'; ExternalWritable := 'False'} : Bool := false;   // Disable step indicated in S_NO
      T_PUSH { ExternalAccessible := 'False'; ExternalVisible := 'False'; ExternalWritable := 'False'} : Bool := false;   // Enable transition to switch in semi automatic mode
      Run : Bool;
      Reset : Bool;
      OwnerIndex : DInt;
      Delta : Time;
   END_VAR
   VAR_OUTPUT
      S_NO { ExternalAccessible := 'False'; ExternalVisible := 'False'; ExternalWritable := 'False'} : Int := 0;   // Step number
      S_MORE { ExternalAccessible := 'False'; ExternalVisible := 'False'; ExternalWritable := 'False'} : Bool := false;   // More steps are available and can be shown in S_NO
      S_ACTIVE { ExternalAccessible := 'False'; ExternalVisible := 'False'; ExternalWritable := 'False'} : Bool := false;   // Step indicated in S_NO is active
      ERR_FLT { ExternalAccessible := 'False'; ExternalVisible := 'False'; ExternalWritable := 'False'} : Bool := false;   // Interlock or supervision group error
      AUTO_ON { ExternalAccessible := 'False'; ExternalVisible := 'False'; ExternalWritable := 'False'} : Bool := false;   // Automatic mode is active
      TAP_ON { ExternalAccessible := 'False'; ExternalVisible := 'False'; ExternalWritable := 'False'} : Bool := false;   // Semiautomatic mode/step with transition enabled
      TOP_ON { ExternalAccessible := 'False'; ExternalVisible := 'False'; ExternalWritable := 'False'} : Bool := false;   // Semiautomatic mode/ignore transition enabled
      MAN_ON { ExternalAccessible := 'False'; ExternalVisible := 'False'; ExternalWritable := 'False'} : Bool := false;   // Manual mode is active
   END_VAR
   VAR_IN_OUT
      PressRam : "FB_CylinderCM";
      Door : "FB_CylinderCM";
      PartSlide : "FB_CylinderCM";
      Seq : "FRK_SequenceCtx";
      Row1 : "FRK_SequenceRow";
      Row2 : "FRK_SequenceRow";
      Row3 : "FRK_SequenceRow";
      Row4 : "FRK_SequenceRow";
      Ready1 { ExternalAccessible := 'False'; ExternalVisible := 'False'; ExternalWritable := 'False'} : Bool;
      Ready2 { ExternalAccessible := 'False'; ExternalVisible := 'False'; ExternalWritable := 'False'} : Bool;
      Ready3 { ExternalAccessible := 'False'; ExternalVisible := 'False'; ExternalWritable := 'False'} : Bool;
      Ready4 { ExternalAccessible := 'False'; ExternalVisible := 'False'; ExternalWritable := 'False'} : Bool;
      Ready5 { ExternalAccessible := 'False'; ExternalVisible := 'False'; ExternalWritable := 'False'} : Bool;
   END_VAR
BEGIN
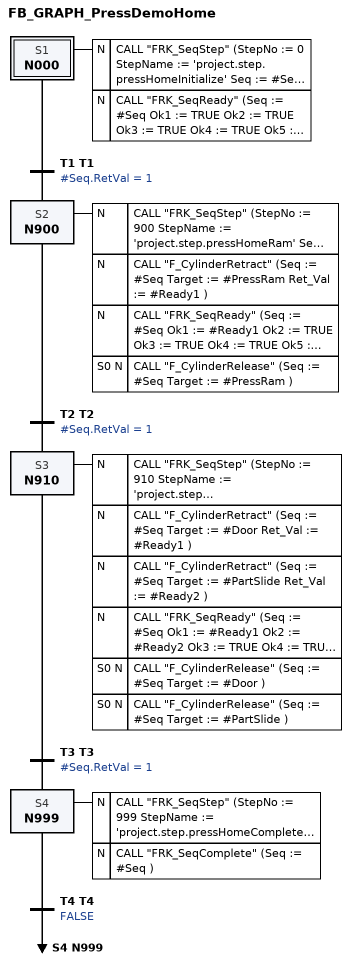
   // sequencer 1
   INITIAL_STEP N000:   // S1, max time T#10S, warning time T#7S
              N    CALL "FRK_SeqStep" 
                   (StepNo := 0
                   StepName := 'project.step.pressHomeInitialize'
                   Seq := #Seq
                   Row := #Row1
                   )
              N    CALL "FRK_SeqReady" 
                   (Seq := #Seq
                   Ok1 := TRUE
                   Ok2 := TRUE
                   Ok3 := TRUE
                   Ok4 := TRUE
                   Ok5 := TRUE
                   )
   END_STEP
   TRANSITION T1 FROM N000 TO N900   // T1
      := #Seq.RetVal = 1;
   END_TRANSITION
   STEP N900:   // S2, max time T#10S, warning time T#7S
              N    CALL "FRK_SeqStep" 
                   (StepNo := 900
                   StepName := 'project.step.pressHomeRam'
                   Seq := #Seq
                   Row := #Row2
                   )
              N    CALL "F_CylinderRetract" 
                   (Seq := #Seq
                   Target := #PressRam
                   Ret_Val := #Ready1
                   )
              N    CALL "FRK_SeqReady" 
                   (Seq := #Seq
                   Ok1 := #Ready1
                   Ok2 := TRUE
                   Ok3 := TRUE
                   Ok4 := TRUE
                   Ok5 := TRUE
                   )
          S0  N    CALL "F_CylinderRelease" 
                   (Seq := #Seq
                   Target := #PressRam
                   )
   END_STEP
   TRANSITION T2 FROM N900 TO N910   // T2
      := #Seq.RetVal = 1;
   END_TRANSITION
   STEP N910:   // S3, max time T#10S, warning time T#7S
              N    CALL "FRK_SeqStep" 
                   (StepNo := 910
                   StepName := 'project.step.pressHomeDoorAndSlide'
                   Seq := #Seq
                   Row := #Row3
                   )
              N    CALL "F_CylinderRetract" 
                   (Seq := #Seq
                   Target := #Door
                   Ret_Val := #Ready1
                   )
              N    CALL "F_CylinderRetract" 
                   (Seq := #Seq
                   Target := #PartSlide
                   Ret_Val := #Ready2
                   )
              N    CALL "FRK_SeqReady" 
                   (Seq := #Seq
                   Ok1 := #Ready1
                   Ok2 := #Ready2
                   Ok3 := TRUE
                   Ok4 := TRUE
                   Ok5 := TRUE
                   )
          S0  N    CALL "F_CylinderRelease" 
                   (Seq := #Seq
                   Target := #Door
                   )
          S0  N    CALL "F_CylinderRelease" 
                   (Seq := #Seq
                   Target := #PartSlide
                   )
   END_STEP
   TRANSITION T3 FROM N910 TO N999   // T3
      := #Seq.RetVal = 1;
   END_TRANSITION
   STEP N999:   // S4, max time T#10S, warning time T#7S
              N    CALL "FRK_SeqStep" 
                   (StepNo := 999
                   StepName := 'project.step.pressHomeComplete'
                   Seq := #Seq
                   Row := #Row4
                   )
              N    CALL "FRK_SeqComplete" 
                   (Seq := #Seq
                   )
   END_STEP
   TRANSITION T4 FROM N999 TO N999   // T4, jump
      := FALSE;
   END_TRANSITION
END_FUNCTION_BLOCK

FUNCTION_BLOCK "FB_LD_PressDemoAuto"   // FB6, LAD
{ S7_Optimized_Access := 'TRUE' }
VERSION : 0.1
// stored: AutoNumber true, IsIECCheckEnabled false, IsRetainMemResEnabled false, MemoryReserve 100, SetENOAutomatically false, UDAEnableTagReadback false
   VAR_INPUT
      Run { ExternalWritable := 'False'} : Bool;
      Reset { ExternalWritable := 'False'} : Bool;
      OwnerIndex { ExternalWritable := 'False'} : DInt;
      Delta { ExternalWritable := 'False'} : Time;
      TransferSettleTime { ExternalWritable := 'False'} : Time;
      PartQuality { ExternalWritable := 'False'} : Bool;
      RequireTwoHandStart { ExternalWritable := 'False'} : Bool;
      SourcePath { ExternalWritable := 'False'} : String[80];
      PartPresent { ExternalWritable := 'False'} : Bool;
      AirPressureOk { ExternalWritable := 'False'} : Bool;
      TwoHandHeld { ExternalWritable := 'False'} : Bool;
      StartPulse { ExternalWritable := 'False'} : Bool;
      PressSettleTime { ExternalWritable := 'False'} : Time;
   END_VAR
   VAR_IN_OUT
      PressRam : "FB_CylinderCM";
      Door : "FB_CylinderCM";
      PartSlide : "FB_CylinderCM";
      Core : "FRK_Core";
      Unit : "FRK_Unit";
      Status : "ST_ModuleStatus";
      Part : "ST_PartContext";
      AlarmLog : "FRK_AlarmLog";
   END_VAR
   VAR
      Seq { ExternalWritable := 'False'} : "FRK_SequenceCtx";
      Row1 { ExternalWritable := 'False'} : "FRK_SequenceRow";
      Row2 { ExternalWritable := 'False'} : "FRK_SequenceRow";
      Row3 { ExternalWritable := 'False'} : "FRK_SequenceRow";
      Row4 { ExternalWritable := 'False'} : "FRK_SequenceRow";
      Row5 { ExternalWritable := 'False'} : "FRK_SequenceRow";
      Row6 { ExternalWritable := 'False'} : "FRK_SequenceRow";
      Row7 { ExternalWritable := 'False'} : "FRK_SequenceRow";
      Row8 { ExternalWritable := 'False'} : "FRK_SequenceRow";
      Row9 { ExternalWritable := 'False'} : "FRK_SequenceRow";
      Row10 { ExternalWritable := 'False'} : "FRK_SequenceRow";
      Row11 { ExternalWritable := 'False'} : "FRK_SequenceRow";
      Row12 { ExternalWritable := 'False'} : "FRK_SequenceRow";
      Row13 { ExternalWritable := 'False'} : "FRK_SequenceRow";
      Row14 { ExternalWritable := 'False'} : "FRK_SequenceRow";
      Row15 { ExternalWritable := 'False'} : "FRK_SequenceRow";
      Row16 { ExternalWritable := 'False'} : "FRK_SequenceRow";
      At0 { ExternalAccessible := 'False'; ExternalVisible := 'False'; ExternalWritable := 'False'} : Bool;
      At100 { ExternalAccessible := 'False'; ExternalVisible := 'False'; ExternalWritable := 'False'} : Bool;
      At110 { ExternalAccessible := 'False'; ExternalVisible := 'False'; ExternalWritable := 'False'} : Bool;
      At130 { ExternalAccessible := 'False'; ExternalVisible := 'False'; ExternalWritable := 'False'} : Bool;
      At150 { ExternalAccessible := 'False'; ExternalVisible := 'False'; ExternalWritable := 'False'} : Bool;
      At170 { ExternalAccessible := 'False'; ExternalVisible := 'False'; ExternalWritable := 'False'} : Bool;
      At180 { ExternalAccessible := 'False'; ExternalVisible := 'False'; ExternalWritable := 'False'} : Bool;
      At185 { ExternalAccessible := 'False'; ExternalVisible := 'False'; ExternalWritable := 'False'} : Bool;
      At190 { ExternalAccessible := 'False'; ExternalVisible := 'False'; ExternalWritable := 'False'} : Bool;
      At200 { ExternalAccessible := 'False'; ExternalVisible := 'False'; ExternalWritable := 'False'} : Bool;
      At210 { ExternalAccessible := 'False'; ExternalVisible := 'False'; ExternalWritable := 'False'} : Bool;
      At215 { ExternalAccessible := 'False'; ExternalVisible := 'False'; ExternalWritable := 'False'} : Bool;
      At220 { ExternalAccessible := 'False'; ExternalVisible := 'False'; ExternalWritable := 'False'} : Bool;
      At230 { ExternalAccessible := 'False'; ExternalVisible := 'False'; ExternalWritable := 'False'} : Bool;
      At240 { ExternalAccessible := 'False'; ExternalVisible := 'False'; ExternalWritable := 'False'} : Bool;
      At999 { ExternalAccessible := 'False'; ExternalVisible := 'False'; ExternalWritable := 'False'} : Bool;
      Ready1 { ExternalAccessible := 'False'; ExternalVisible := 'False'; ExternalWritable := 'False'} : Bool;
      Ready2 { ExternalAccessible := 'False'; ExternalVisible := 'False'; ExternalWritable := 'False'} : Bool;
      Ready3 { ExternalAccessible := 'False'; ExternalVisible := 'False'; ExternalWritable := 'False'} : Bool;
      Ready4 { ExternalAccessible := 'False'; ExternalVisible := 'False'; ExternalWritable := 'False'} : Bool;
      Ready5 { ExternalAccessible := 'False'; ExternalVisible := 'False'; ExternalWritable := 'False'} : Bool;
      Advance { ExternalAccessible := 'False'; ExternalVisible := 'False'; ExternalWritable := 'False'} : Bool;
      Cycle { ExternalAccessible := 'False'; ExternalVisible := 'False'; ExternalWritable := 'False'} : "ST_PressDemoCycle";
      LoadPosition { ExternalAccessible := 'False'; ExternalVisible := 'False'; ExternalWritable := 'False'} : "FB_PressDemoLoadPosition";
      LoadDone { ExternalAccessible := 'False'; ExternalVisible := 'False'; ExternalWritable := 'False'} : Bool;
      LoadActive { ExternalAccessible := 'False'; ExternalVisible := 'False'; ExternalWritable := 'False'} : Bool;
   END_VAR
BEGIN

REGION Network 1
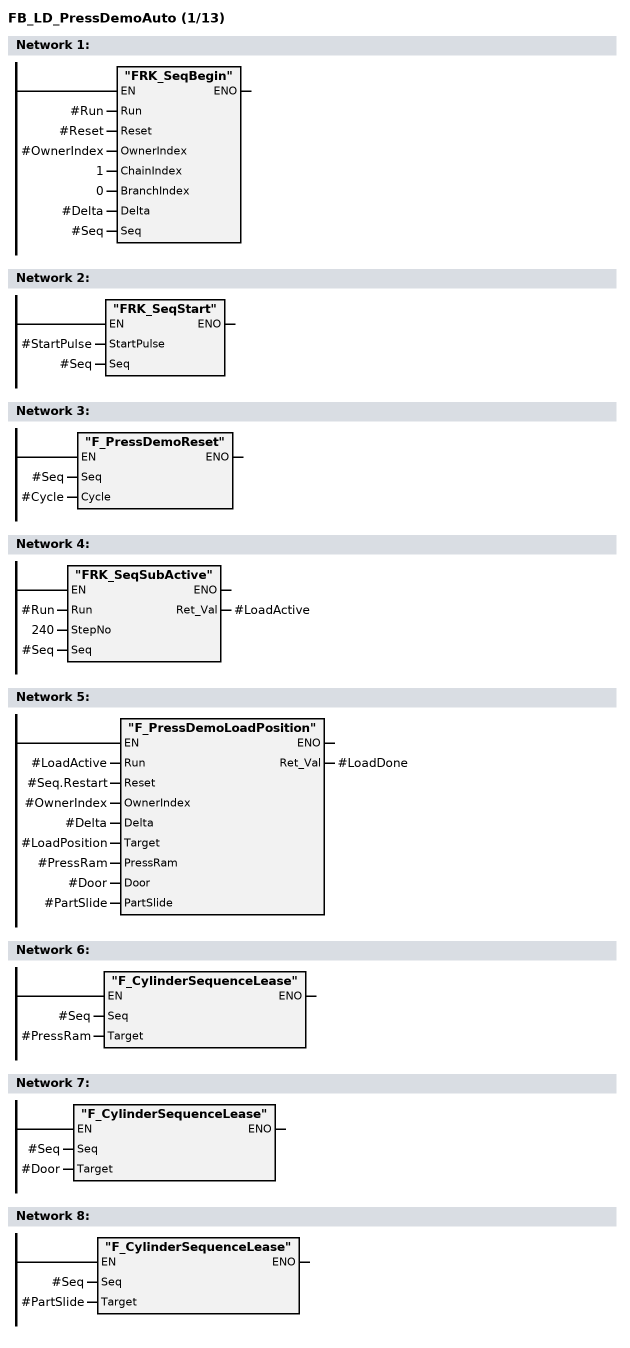
   RUNG wire#powerrail
      "FRK_SeqBegin"(Run := #Run, Reset := #Reset, OwnerIndex := #OwnerIndex, ChainIndex := 1, BranchIndex := 0, Delta := #Delta, Seq := #Seq)
   END_RUNG
   // the same network as SCL:
   "FRK_SeqBegin"(Run := #Run,
                  Reset := #Reset,
                  OwnerIndex := #OwnerIndex,
                  ChainIndex := 1,
                  BranchIndex := 0,
                  Delta := #Delta,
                  Seq := #Seq);
END_REGION

REGION Network 2
   RUNG wire#powerrail
      "FRK_SeqStart"(StartPulse := #StartPulse, Seq := #Seq)
   END_RUNG
   // the same network as SCL:
   "FRK_SeqStart"(StartPulse := #StartPulse, Seq := #Seq);
END_REGION

REGION Network 3
   RUNG wire#powerrail
      "F_PressDemoReset"(Seq := #Seq, Cycle := #Cycle)
   END_RUNG
   // the same network as SCL:
   "F_PressDemoReset"(Seq := #Seq, Cycle := #Cycle);
END_REGION

REGION Network 4
   RUNG wire#powerrail
      "FRK_SeqSubActive"(Run := #Run, StepNo := 240, Seq := #Seq, Ret_Val => #LoadActive)
   END_RUNG
   // the same network as SCL:
   #LoadActive := "FRK_SeqSubActive"(Run := #Run, StepNo := 240, Seq := #Seq);
END_REGION

REGION Network 5
   RUNG wire#powerrail
      "F_PressDemoLoadPosition"(Run := #LoadActive, Reset := #Seq.Restart, OwnerIndex := #OwnerIndex, Delta := #Delta, Target := #LoadPosition, PressRam := #PressRam, Door := #Door, PartSlide := #PartSlide, Ret_Val => #LoadDone)
   END_RUNG
   // the same network as SCL:
   #LoadDone := "F_PressDemoLoadPosition"(Run := #LoadActive,
                           Reset := #Seq.Restart,
                           OwnerIndex := #OwnerIndex,
                           Delta := #Delta,
                           Target := #LoadPosition,
                           PressRam := #PressRam,
                           Door := #Door,
                           PartSlide := #PartSlide);
END_REGION

REGION Network 6
   RUNG wire#powerrail
      "F_CylinderSequenceLease"(Seq := #Seq, Target := #PressRam)
   END_RUNG
   // the same network as SCL:
   "F_CylinderSequenceLease"(Seq := #Seq, Target := #PressRam);
END_REGION

REGION Network 7
   RUNG wire#powerrail
      "F_CylinderSequenceLease"(Seq := #Seq, Target := #Door)
   END_RUNG
   // the same network as SCL:
   "F_CylinderSequenceLease"(Seq := #Seq, Target := #Door);
END_REGION

REGION Network 8
   RUNG wire#powerrail
      "F_CylinderSequenceLease"(Seq := #Seq, Target := #PartSlide)
   END_RUNG
   // the same network as SCL:
   "F_CylinderSequenceLease"(Seq := #Seq, Target := #PartSlide);
END_REGION

REGION Network 9
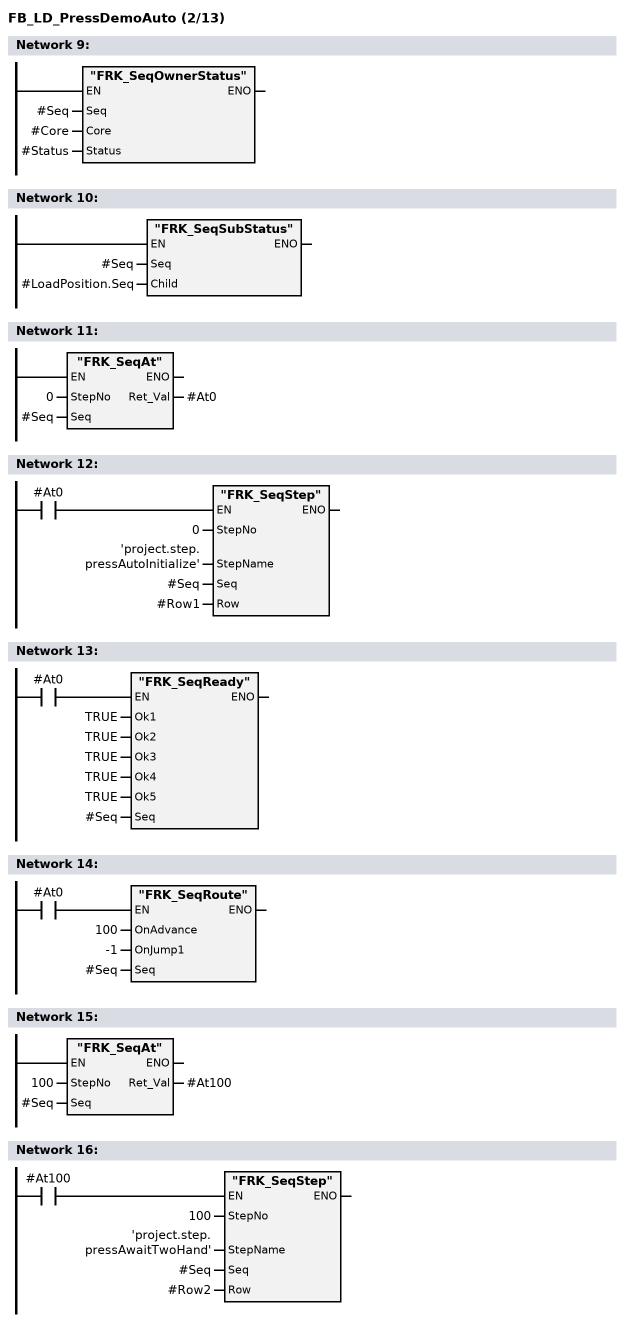
   RUNG wire#powerrail
      "FRK_SeqOwnerStatus"(Seq := #Seq, Core := #Core, Status := #Status)
   END_RUNG
   // the same network as SCL:
   "FRK_SeqOwnerStatus"(Seq := #Seq, Core := #Core, Status := #Status);
END_REGION

REGION Network 10
   RUNG wire#powerrail
      "FRK_SeqSubStatus"(Seq := #Seq, Child := #LoadPosition.Seq)
   END_RUNG
   // the same network as SCL:
   "FRK_SeqSubStatus"(Seq := #Seq, Child := #LoadPosition.Seq);
END_REGION

REGION Network 11
   RUNG wire#powerrail
      "FRK_SeqAt"(StepNo := 0, Seq := #Seq, Ret_Val => #At0)
   END_RUNG
   // the same network as SCL:
   #At0 := "FRK_SeqAt"(StepNo := 0, Seq := #Seq);
END_REGION

REGION Network 12
   RUNG wire#powerrail
      Contact( #At0 )
      "FRK_SeqStep"(StepNo := 0, StepName := 'project.step.pressAutoInitialize', Seq := #Seq, Row := #Row1)
   END_RUNG
   // the same network as SCL:
   IF #At0 THEN
       "FRK_SeqStep"(StepNo := 0, StepName := 'project.step.pressAutoInitialize', Seq := #Seq, Row := #Row1);
   END_IF;
END_REGION

REGION Network 13
   RUNG wire#powerrail
      Contact( #At0 )
      "FRK_SeqReady"(Ok1 := TRUE, Ok2 := TRUE, Ok3 := TRUE, Ok4 := TRUE, Ok5 := TRUE, Seq := #Seq)
   END_RUNG
   // the same network as SCL:
   IF #At0 THEN
       "FRK_SeqReady"(Ok1 := TRUE, Ok2 := TRUE, Ok3 := TRUE, Ok4 := TRUE, Ok5 := TRUE, Seq := #Seq);
   END_IF;
END_REGION

REGION Network 14
   RUNG wire#powerrail
      Contact( #At0 )
      "FRK_SeqRoute"(OnAdvance := 100, OnJump1 := -1, Seq := #Seq)
   END_RUNG
   // the same network as SCL:
   IF #At0 THEN "FRK_SeqRoute"(OnAdvance := 100, OnJump1 := -1, Seq := #Seq); END_IF;
END_REGION

REGION Network 15
   RUNG wire#powerrail
      "FRK_SeqAt"(StepNo := 100, Seq := #Seq, Ret_Val => #At100)
   END_RUNG
   // the same network as SCL:
   #At100 := "FRK_SeqAt"(StepNo := 100, Seq := #Seq);
END_REGION

REGION Network 16
   RUNG wire#powerrail
      Contact( #At100 )
      "FRK_SeqStep"(StepNo := 100, StepName := 'project.step.pressAwaitTwoHand', Seq := #Seq, Row := #Row2)
   END_RUNG
   // the same network as SCL:
   IF #At100 THEN
       "FRK_SeqStep"(StepNo := 100, StepName := 'project.step.pressAwaitTwoHand', Seq := #Seq, Row := #Row2);
   END_IF;
END_REGION

REGION Network 17
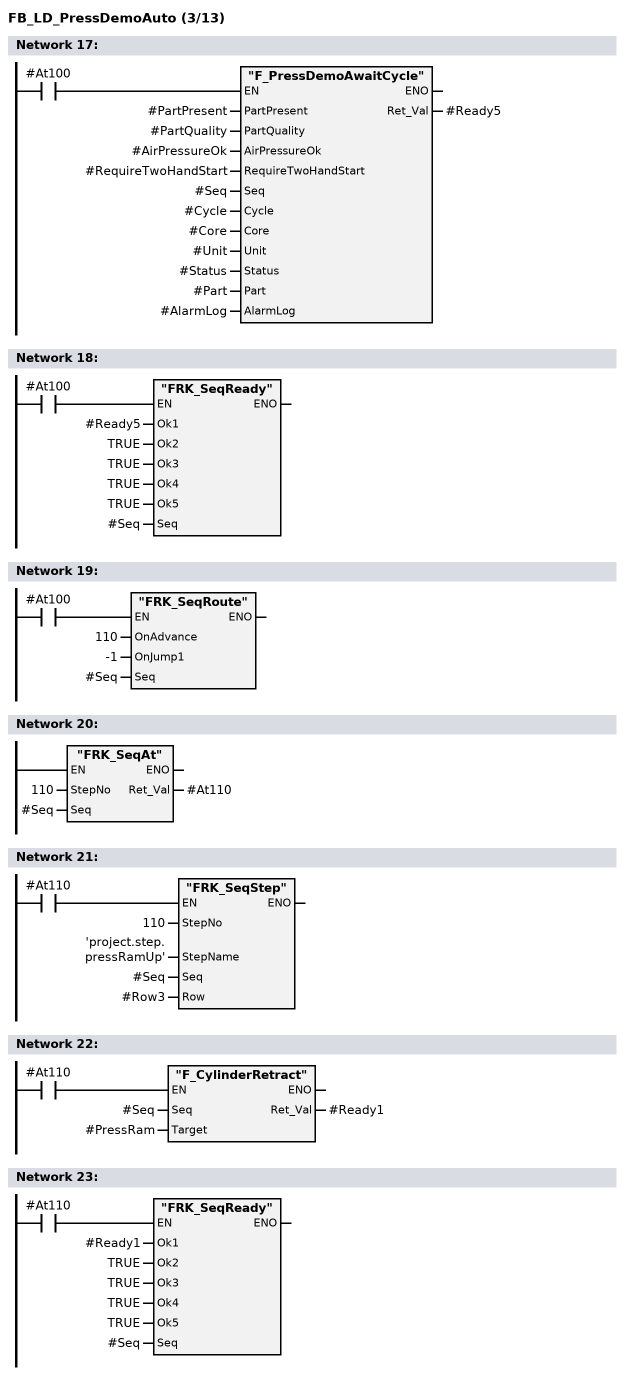
   RUNG wire#powerrail
      Contact( #At100 )
      "F_PressDemoAwaitCycle"(PartPresent := #PartPresent, PartQuality := #PartQuality, AirPressureOk := #AirPressureOk, RequireTwoHandStart := #RequireTwoHandStart, Seq := #Seq, Cycle := #Cycle, Core := #Core, Unit := #Unit, Status := #Status, Part := #Part, AlarmLog := #AlarmLog, Ret_Val => #Ready5)
   END_RUNG
   // the same network as SCL:
   IF #At100 THEN
       #Ready5 := "F_PressDemoAwaitCycle"(PartPresent := #PartPresent,
                               PartQuality := #PartQuality,
                               AirPressureOk := #AirPressureOk,
                               RequireTwoHandStart := #RequireTwoHandStart,
                               Seq := #Seq,
                               Cycle := #Cycle,
                               Core := #Core,
                               Unit := #Unit,
                               Status := #Status,
                               Part := #Part,
                               AlarmLog := #AlarmLog);
   END_IF;
END_REGION

REGION Network 18
   RUNG wire#powerrail
      Contact( #At100 )
      "FRK_SeqReady"(Ok1 := #Ready5, Ok2 := TRUE, Ok3 := TRUE, Ok4 := TRUE, Ok5 := TRUE, Seq := #Seq)
   END_RUNG
   // the same network as SCL:
   IF #At100 THEN
       "FRK_SeqReady"(Ok1 := #Ready5, Ok2 := TRUE, Ok3 := TRUE, Ok4 := TRUE, Ok5 := TRUE, Seq := #Seq);
   END_IF;
END_REGION

REGION Network 19
   RUNG wire#powerrail
      Contact( #At100 )
      "FRK_SeqRoute"(OnAdvance := 110, OnJump1 := -1, Seq := #Seq)
   END_RUNG
   // the same network as SCL:
   IF #At100 THEN "FRK_SeqRoute"(OnAdvance := 110, OnJump1 := -1, Seq := #Seq); END_IF;
END_REGION

REGION Network 20
   RUNG wire#powerrail
      "FRK_SeqAt"(StepNo := 110, Seq := #Seq, Ret_Val => #At110)
   END_RUNG
   // the same network as SCL:
   #At110 := "FRK_SeqAt"(StepNo := 110, Seq := #Seq);
END_REGION

REGION Network 21
   RUNG wire#powerrail
      Contact( #At110 )
      "FRK_SeqStep"(StepNo := 110, StepName := 'project.step.pressRamUp', Seq := #Seq, Row := #Row3)
   END_RUNG
   // the same network as SCL:
   IF #At110 THEN
       "FRK_SeqStep"(StepNo := 110, StepName := 'project.step.pressRamUp', Seq := #Seq, Row := #Row3);
   END_IF;
END_REGION

REGION Network 22
   RUNG wire#powerrail
      Contact( #At110 )
      "F_CylinderRetract"(Seq := #Seq, Target := #PressRam, Ret_Val => #Ready1)
   END_RUNG
   // the same network as SCL:
   IF #At110 THEN #Ready1 := "F_CylinderRetract"(Seq := #Seq, Target := #PressRam); END_IF;
END_REGION

REGION Network 23
   RUNG wire#powerrail
      Contact( #At110 )
      "FRK_SeqReady"(Ok1 := #Ready1, Ok2 := TRUE, Ok3 := TRUE, Ok4 := TRUE, Ok5 := TRUE, Seq := #Seq)
   END_RUNG
   // the same network as SCL:
   IF #At110 THEN
       "FRK_SeqReady"(Ok1 := #Ready1, Ok2 := TRUE, Ok3 := TRUE, Ok4 := TRUE, Ok5 := TRUE, Seq := #Seq);
   END_IF;
END_REGION

REGION Network 24
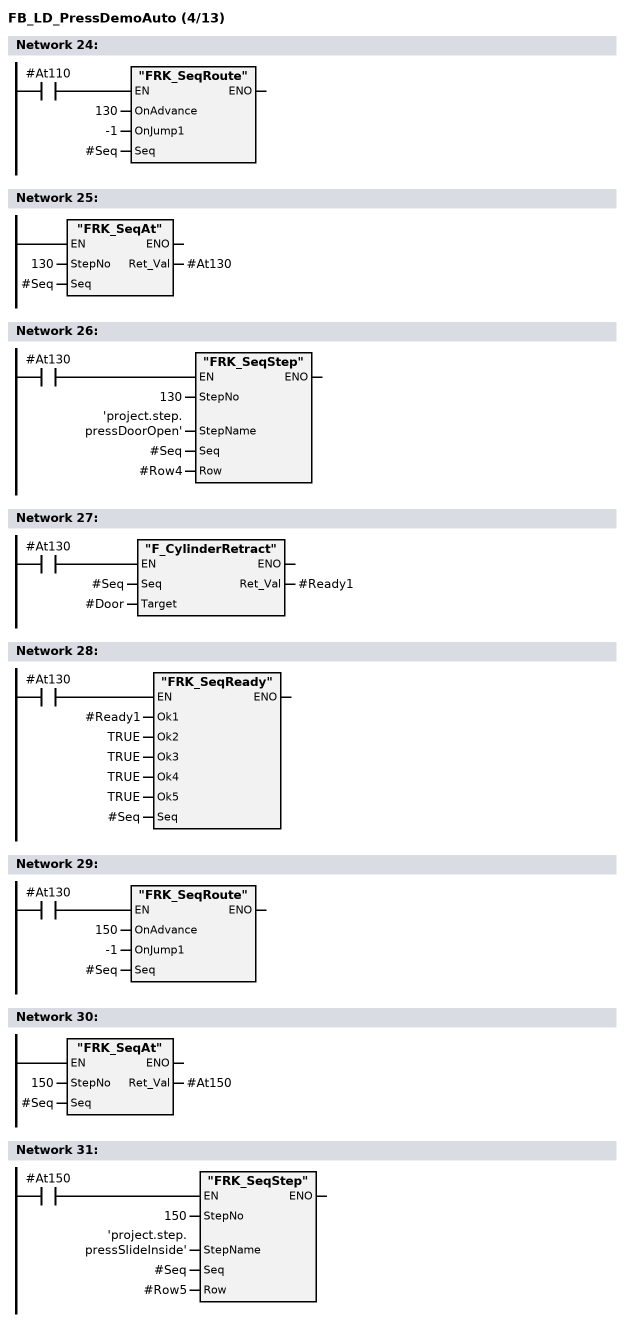
   RUNG wire#powerrail
      Contact( #At110 )
      "FRK_SeqRoute"(OnAdvance := 130, OnJump1 := -1, Seq := #Seq)
   END_RUNG
   // the same network as SCL:
   IF #At110 THEN "FRK_SeqRoute"(OnAdvance := 130, OnJump1 := -1, Seq := #Seq); END_IF;
END_REGION

REGION Network 25
   RUNG wire#powerrail
      "FRK_SeqAt"(StepNo := 130, Seq := #Seq, Ret_Val => #At130)
   END_RUNG
   // the same network as SCL:
   #At130 := "FRK_SeqAt"(StepNo := 130, Seq := #Seq);
END_REGION

REGION Network 26
   RUNG wire#powerrail
      Contact( #At130 )
      "FRK_SeqStep"(StepNo := 130, StepName := 'project.step.pressDoorOpen', Seq := #Seq, Row := #Row4)
   END_RUNG
   // the same network as SCL:
   IF #At130 THEN
       "FRK_SeqStep"(StepNo := 130, StepName := 'project.step.pressDoorOpen', Seq := #Seq, Row := #Row4);
   END_IF;
END_REGION

REGION Network 27
   RUNG wire#powerrail
      Contact( #At130 )
      "F_CylinderRetract"(Seq := #Seq, Target := #Door, Ret_Val => #Ready1)
   END_RUNG
   // the same network as SCL:
   IF #At130 THEN #Ready1 := "F_CylinderRetract"(Seq := #Seq, Target := #Door); END_IF;
END_REGION

REGION Network 28
   RUNG wire#powerrail
      Contact( #At130 )
      "FRK_SeqReady"(Ok1 := #Ready1, Ok2 := TRUE, Ok3 := TRUE, Ok4 := TRUE, Ok5 := TRUE, Seq := #Seq)
   END_RUNG
   // the same network as SCL:
   IF #At130 THEN
       "FRK_SeqReady"(Ok1 := #Ready1, Ok2 := TRUE, Ok3 := TRUE, Ok4 := TRUE, Ok5 := TRUE, Seq := #Seq);
   END_IF;
END_REGION

REGION Network 29
   RUNG wire#powerrail
      Contact( #At130 )
      "FRK_SeqRoute"(OnAdvance := 150, OnJump1 := -1, Seq := #Seq)
   END_RUNG
   // the same network as SCL:
   IF #At130 THEN "FRK_SeqRoute"(OnAdvance := 150, OnJump1 := -1, Seq := #Seq); END_IF;
END_REGION

REGION Network 30
   RUNG wire#powerrail
      "FRK_SeqAt"(StepNo := 150, Seq := #Seq, Ret_Val => #At150)
   END_RUNG
   // the same network as SCL:
   #At150 := "FRK_SeqAt"(StepNo := 150, Seq := #Seq);
END_REGION

REGION Network 31
   RUNG wire#powerrail
      Contact( #At150 )
      "FRK_SeqStep"(StepNo := 150, StepName := 'project.step.pressSlideInside', Seq := #Seq, Row := #Row5)
   END_RUNG
   // the same network as SCL:
   IF #At150 THEN
       "FRK_SeqStep"(StepNo := 150, StepName := 'project.step.pressSlideInside', Seq := #Seq, Row := #Row5);
   END_IF;
END_REGION

REGION Network 32
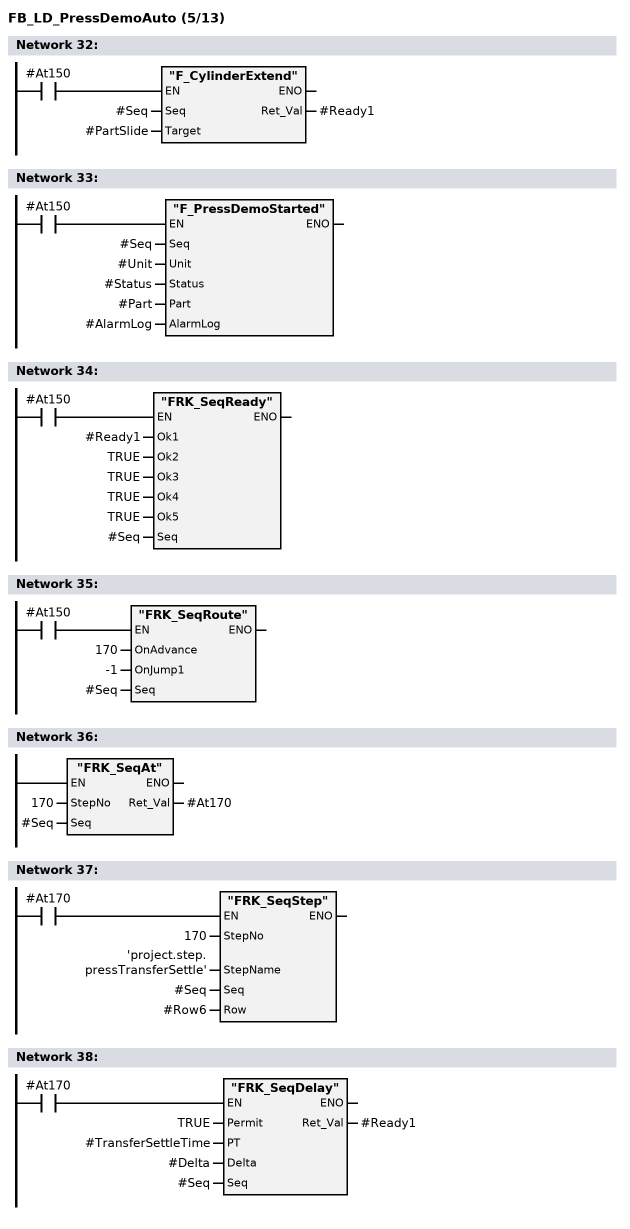
   RUNG wire#powerrail
      Contact( #At150 )
      "F_CylinderExtend"(Seq := #Seq, Target := #PartSlide, Ret_Val => #Ready1)
   END_RUNG
   // the same network as SCL:
   IF #At150 THEN #Ready1 := "F_CylinderExtend"(Seq := #Seq, Target := #PartSlide); END_IF;
END_REGION

REGION Network 33
   RUNG wire#powerrail
      Contact( #At150 )
      "F_PressDemoStarted"(Seq := #Seq, Unit := #Unit, Status := #Status, Part := #Part, AlarmLog := #AlarmLog)
   END_RUNG
   // the same network as SCL:
   IF #At150 THEN
       "F_PressDemoStarted"(Seq := #Seq, Unit := #Unit, Status := #Status, Part := #Part, AlarmLog := #AlarmLog);
   END_IF;
END_REGION

REGION Network 34
   RUNG wire#powerrail
      Contact( #At150 )
      "FRK_SeqReady"(Ok1 := #Ready1, Ok2 := TRUE, Ok3 := TRUE, Ok4 := TRUE, Ok5 := TRUE, Seq := #Seq)
   END_RUNG
   // the same network as SCL:
   IF #At150 THEN
       "FRK_SeqReady"(Ok1 := #Ready1, Ok2 := TRUE, Ok3 := TRUE, Ok4 := TRUE, Ok5 := TRUE, Seq := #Seq);
   END_IF;
END_REGION

REGION Network 35
   RUNG wire#powerrail
      Contact( #At150 )
      "FRK_SeqRoute"(OnAdvance := 170, OnJump1 := -1, Seq := #Seq)
   END_RUNG
   // the same network as SCL:
   IF #At150 THEN "FRK_SeqRoute"(OnAdvance := 170, OnJump1 := -1, Seq := #Seq); END_IF;
END_REGION

REGION Network 36
   RUNG wire#powerrail
      "FRK_SeqAt"(StepNo := 170, Seq := #Seq, Ret_Val => #At170)
   END_RUNG
   // the same network as SCL:
   #At170 := "FRK_SeqAt"(StepNo := 170, Seq := #Seq);
END_REGION

REGION Network 37
   RUNG wire#powerrail
      Contact( #At170 )
      "FRK_SeqStep"(StepNo := 170, StepName := 'project.step.pressTransferSettle', Seq := #Seq, Row := #Row6)
   END_RUNG
   // the same network as SCL:
   IF #At170 THEN
       "FRK_SeqStep"(StepNo := 170, StepName := 'project.step.pressTransferSettle', Seq := #Seq, Row := #Row6);
   END_IF;
END_REGION

REGION Network 38
   RUNG wire#powerrail
      Contact( #At170 )
      "FRK_SeqDelay"(Permit := TRUE, PT := #TransferSettleTime, Delta := #Delta, Seq := #Seq, Ret_Val => #Ready1)
   END_RUNG
   // the same network as SCL:
   IF #At170 THEN
       #Ready1 := "FRK_SeqDelay"(Permit := TRUE, PT := #TransferSettleTime, Delta := #Delta, Seq := #Seq);
   END_IF;
END_REGION

REGION Network 39
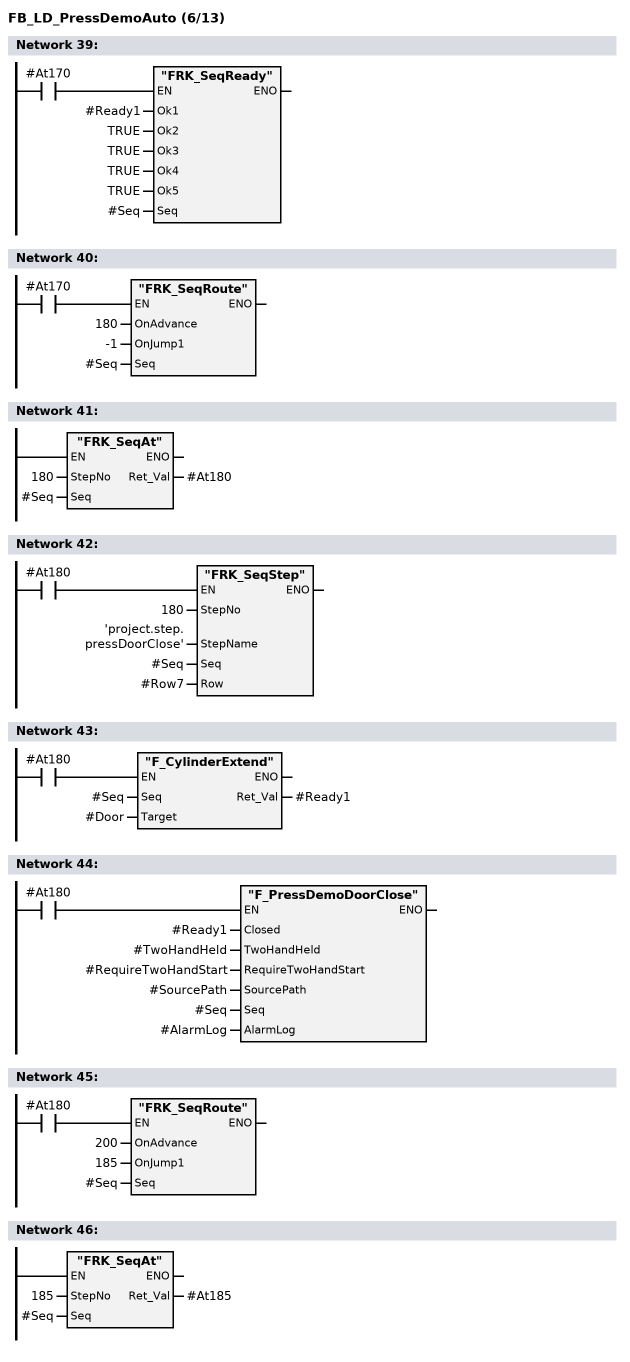
   RUNG wire#powerrail
      Contact( #At170 )
      "FRK_SeqReady"(Ok1 := #Ready1, Ok2 := TRUE, Ok3 := TRUE, Ok4 := TRUE, Ok5 := TRUE, Seq := #Seq)
   END_RUNG
   // the same network as SCL:
   IF #At170 THEN
       "FRK_SeqReady"(Ok1 := #Ready1, Ok2 := TRUE, Ok3 := TRUE, Ok4 := TRUE, Ok5 := TRUE, Seq := #Seq);
   END_IF;
END_REGION

REGION Network 40
   RUNG wire#powerrail
      Contact( #At170 )
      "FRK_SeqRoute"(OnAdvance := 180, OnJump1 := -1, Seq := #Seq)
   END_RUNG
   // the same network as SCL:
   IF #At170 THEN "FRK_SeqRoute"(OnAdvance := 180, OnJump1 := -1, Seq := #Seq); END_IF;
END_REGION

REGION Network 41
   RUNG wire#powerrail
      "FRK_SeqAt"(StepNo := 180, Seq := #Seq, Ret_Val => #At180)
   END_RUNG
   // the same network as SCL:
   #At180 := "FRK_SeqAt"(StepNo := 180, Seq := #Seq);
END_REGION

REGION Network 42
   RUNG wire#powerrail
      Contact( #At180 )
      "FRK_SeqStep"(StepNo := 180, StepName := 'project.step.pressDoorClose', Seq := #Seq, Row := #Row7)
   END_RUNG
   // the same network as SCL:
   IF #At180 THEN
       "FRK_SeqStep"(StepNo := 180, StepName := 'project.step.pressDoorClose', Seq := #Seq, Row := #Row7);
   END_IF;
END_REGION

REGION Network 43
   RUNG wire#powerrail
      Contact( #At180 )
      "F_CylinderExtend"(Seq := #Seq, Target := #Door, Ret_Val => #Ready1)
   END_RUNG
   // the same network as SCL:
   IF #At180 THEN #Ready1 := "F_CylinderExtend"(Seq := #Seq, Target := #Door); END_IF;
END_REGION

REGION Network 44
   RUNG wire#powerrail
      Contact( #At180 )
      "F_PressDemoDoorClose"(Closed := #Ready1, TwoHandHeld := #TwoHandHeld, RequireTwoHandStart := #RequireTwoHandStart, SourcePath := #SourcePath, Seq := #Seq, AlarmLog := #AlarmLog)
   END_RUNG
   // the same network as SCL:
   IF #At180 THEN
       "F_PressDemoDoorClose"(Closed := #Ready1,
                              TwoHandHeld := #TwoHandHeld,
                              RequireTwoHandStart := #RequireTwoHandStart,
                              SourcePath := #SourcePath,
                              Seq := #Seq,
                              AlarmLog := #AlarmLog);
   END_IF;
END_REGION

REGION Network 45
   RUNG wire#powerrail
      Contact( #At180 )
      "FRK_SeqRoute"(OnAdvance := 200, OnJump1 := 185, Seq := #Seq)
   END_RUNG
   // the same network as SCL:
   IF #At180 THEN "FRK_SeqRoute"(OnAdvance := 200, OnJump1 := 185, Seq := #Seq); END_IF;
END_REGION

REGION Network 46
   RUNG wire#powerrail
      "FRK_SeqAt"(StepNo := 185, Seq := #Seq, Ret_Val => #At185)
   END_RUNG
   // the same network as SCL:
   #At185 := "FRK_SeqAt"(StepNo := 185, Seq := #Seq);
END_REGION

REGION Network 47
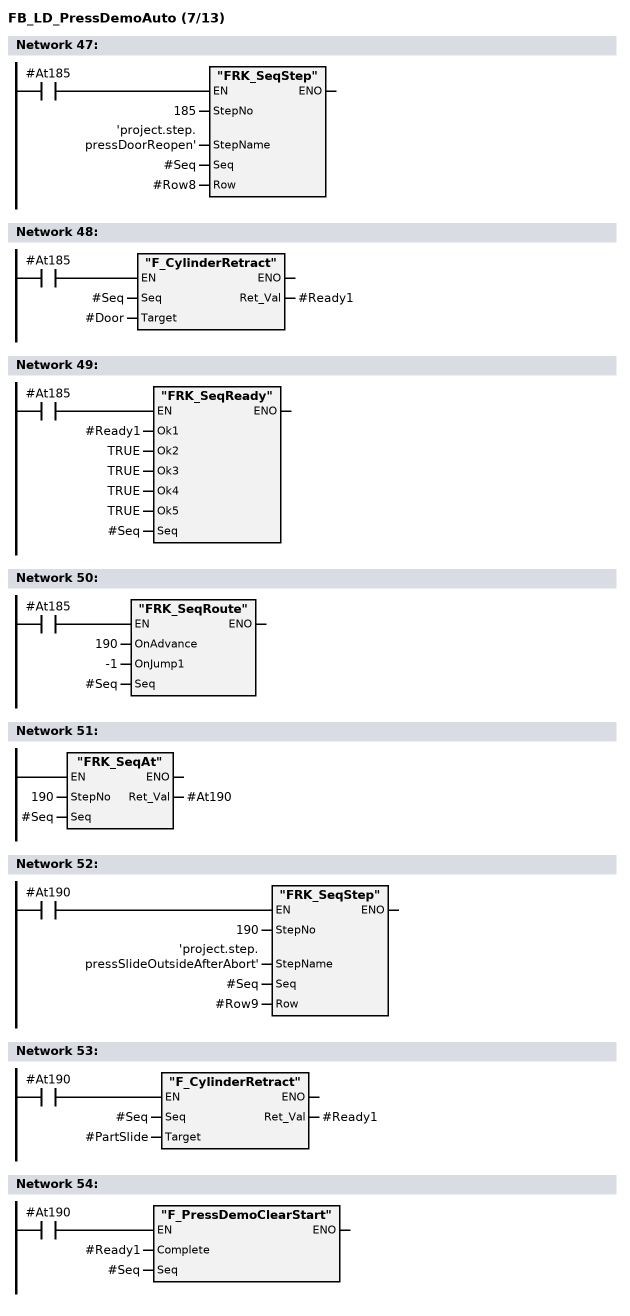
   RUNG wire#powerrail
      Contact( #At185 )
      "FRK_SeqStep"(StepNo := 185, StepName := 'project.step.pressDoorReopen', Seq := #Seq, Row := #Row8)
   END_RUNG
   // the same network as SCL:
   IF #At185 THEN
       "FRK_SeqStep"(StepNo := 185, StepName := 'project.step.pressDoorReopen', Seq := #Seq, Row := #Row8);
   END_IF;
END_REGION

REGION Network 48
   RUNG wire#powerrail
      Contact( #At185 )
      "F_CylinderRetract"(Seq := #Seq, Target := #Door, Ret_Val => #Ready1)
   END_RUNG
   // the same network as SCL:
   IF #At185 THEN #Ready1 := "F_CylinderRetract"(Seq := #Seq, Target := #Door); END_IF;
END_REGION

REGION Network 49
   RUNG wire#powerrail
      Contact( #At185 )
      "FRK_SeqReady"(Ok1 := #Ready1, Ok2 := TRUE, Ok3 := TRUE, Ok4 := TRUE, Ok5 := TRUE, Seq := #Seq)
   END_RUNG
   // the same network as SCL:
   IF #At185 THEN
       "FRK_SeqReady"(Ok1 := #Ready1, Ok2 := TRUE, Ok3 := TRUE, Ok4 := TRUE, Ok5 := TRUE, Seq := #Seq);
   END_IF;
END_REGION

REGION Network 50
   RUNG wire#powerrail
      Contact( #At185 )
      "FRK_SeqRoute"(OnAdvance := 190, OnJump1 := -1, Seq := #Seq)
   END_RUNG
   // the same network as SCL:
   IF #At185 THEN "FRK_SeqRoute"(OnAdvance := 190, OnJump1 := -1, Seq := #Seq); END_IF;
END_REGION

REGION Network 51
   RUNG wire#powerrail
      "FRK_SeqAt"(StepNo := 190, Seq := #Seq, Ret_Val => #At190)
   END_RUNG
   // the same network as SCL:
   #At190 := "FRK_SeqAt"(StepNo := 190, Seq := #Seq);
END_REGION

REGION Network 52
   RUNG wire#powerrail
      Contact( #At190 )
      "FRK_SeqStep"(StepNo := 190, StepName := 'project.step.pressSlideOutsideAfterAbort', Seq := #Seq, Row := #Row9)
   END_RUNG
   // the same network as SCL:
   IF #At190 THEN
       "FRK_SeqStep"(StepNo := 190,
                     StepName := 'project.step.pressSlideOutsideAfterAbort',
                     Seq := #Seq,
                     Row := #Row9);
   END_IF;
END_REGION

REGION Network 53
   RUNG wire#powerrail
      Contact( #At190 )
      "F_CylinderRetract"(Seq := #Seq, Target := #PartSlide, Ret_Val => #Ready1)
   END_RUNG
   // the same network as SCL:
   IF #At190 THEN #Ready1 := "F_CylinderRetract"(Seq := #Seq, Target := #PartSlide); END_IF;
END_REGION

REGION Network 54
   RUNG wire#powerrail
      Contact( #At190 )
      "F_PressDemoClearStart"(Complete := #Ready1, Seq := #Seq)
   END_RUNG
   // the same network as SCL:
   IF #At190 THEN "F_PressDemoClearStart"(Complete := #Ready1, Seq := #Seq); END_IF;
END_REGION

REGION Network 55
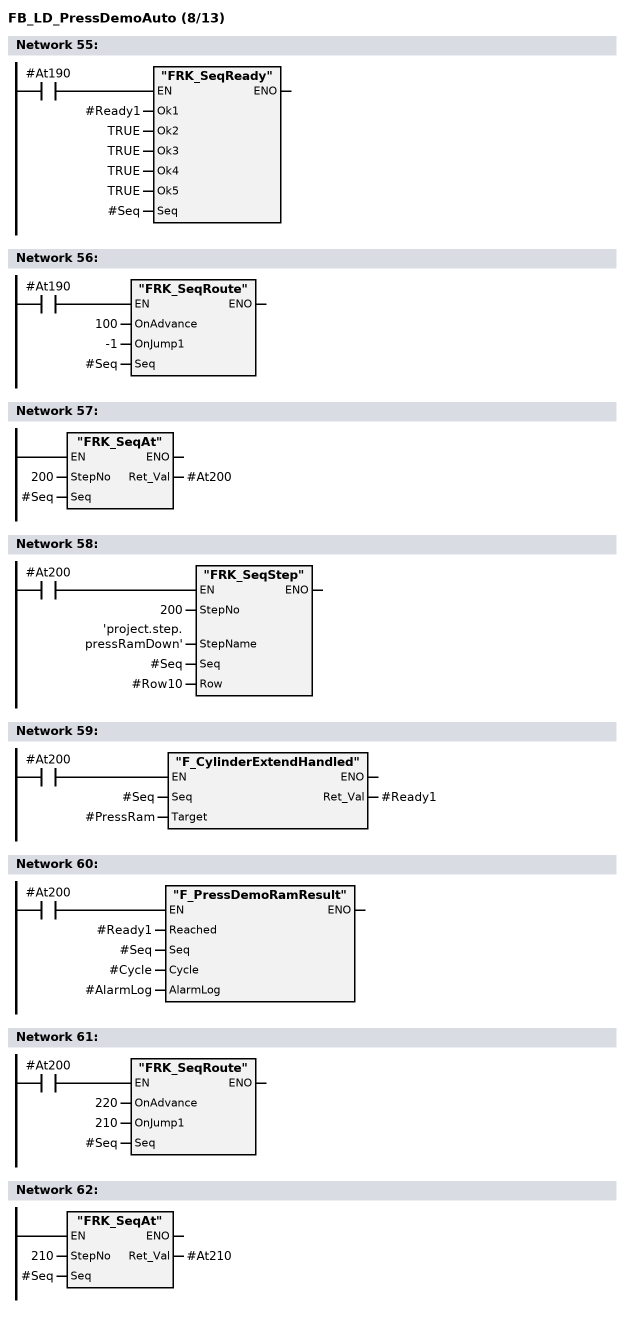
   RUNG wire#powerrail
      Contact( #At190 )
      "FRK_SeqReady"(Ok1 := #Ready1, Ok2 := TRUE, Ok3 := TRUE, Ok4 := TRUE, Ok5 := TRUE, Seq := #Seq)
   END_RUNG
   // the same network as SCL:
   IF #At190 THEN
       "FRK_SeqReady"(Ok1 := #Ready1, Ok2 := TRUE, Ok3 := TRUE, Ok4 := TRUE, Ok5 := TRUE, Seq := #Seq);
   END_IF;
END_REGION

REGION Network 56
   RUNG wire#powerrail
      Contact( #At190 )
      "FRK_SeqRoute"(OnAdvance := 100, OnJump1 := -1, Seq := #Seq)
   END_RUNG
   // the same network as SCL:
   IF #At190 THEN "FRK_SeqRoute"(OnAdvance := 100, OnJump1 := -1, Seq := #Seq); END_IF;
END_REGION

REGION Network 57
   RUNG wire#powerrail
      "FRK_SeqAt"(StepNo := 200, Seq := #Seq, Ret_Val => #At200)
   END_RUNG
   // the same network as SCL:
   #At200 := "FRK_SeqAt"(StepNo := 200, Seq := #Seq);
END_REGION

REGION Network 58
   RUNG wire#powerrail
      Contact( #At200 )
      "FRK_SeqStep"(StepNo := 200, StepName := 'project.step.pressRamDown', Seq := #Seq, Row := #Row10)
   END_RUNG
   // the same network as SCL:
   IF #At200 THEN
       "FRK_SeqStep"(StepNo := 200, StepName := 'project.step.pressRamDown', Seq := #Seq, Row := #Row10);
   END_IF;
END_REGION

REGION Network 59
   RUNG wire#powerrail
      Contact( #At200 )
      "F_CylinderExtendHandled"(Seq := #Seq, Target := #PressRam, Ret_Val => #Ready1)
   END_RUNG
   // the same network as SCL:
   IF #At200 THEN #Ready1 := "F_CylinderExtendHandled"(Seq := #Seq, Target := #PressRam); END_IF;
END_REGION

REGION Network 60
   RUNG wire#powerrail
      Contact( #At200 )
      "F_PressDemoRamResult"(Reached := #Ready1, Seq := #Seq, Cycle := #Cycle, AlarmLog := #AlarmLog)
   END_RUNG
   // the same network as SCL:
   IF #At200 THEN
       "F_PressDemoRamResult"(Reached := #Ready1, Seq := #Seq, Cycle := #Cycle, AlarmLog := #AlarmLog);
   END_IF;
END_REGION

REGION Network 61
   RUNG wire#powerrail
      Contact( #At200 )
      "FRK_SeqRoute"(OnAdvance := 220, OnJump1 := 210, Seq := #Seq)
   END_RUNG
   // the same network as SCL:
   IF #At200 THEN "FRK_SeqRoute"(OnAdvance := 220, OnJump1 := 210, Seq := #Seq); END_IF;
END_REGION

REGION Network 62
   RUNG wire#powerrail
      "FRK_SeqAt"(StepNo := 210, Seq := #Seq, Ret_Val => #At210)
   END_RUNG
   // the same network as SCL:
   #At210 := "FRK_SeqAt"(StepNo := 210, Seq := #Seq);
END_REGION

REGION Network 63
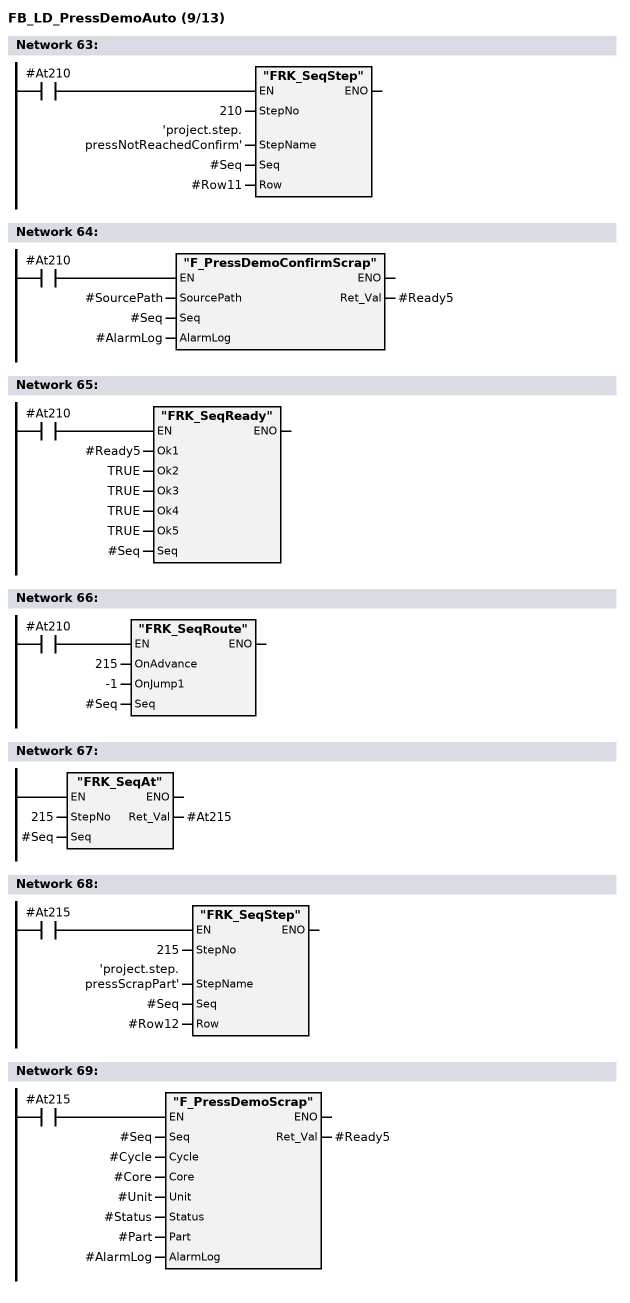
   RUNG wire#powerrail
      Contact( #At210 )
      "FRK_SeqStep"(StepNo := 210, StepName := 'project.step.pressNotReachedConfirm', Seq := #Seq, Row := #Row11)
   END_RUNG
   // the same network as SCL:
   IF #At210 THEN
       "FRK_SeqStep"(StepNo := 210, StepName := 'project.step.pressNotReachedConfirm', Seq := #Seq, Row := #Row11);
   END_IF;
END_REGION

REGION Network 64
   RUNG wire#powerrail
      Contact( #At210 )
      "F_PressDemoConfirmScrap"(SourcePath := #SourcePath, Seq := #Seq, AlarmLog := #AlarmLog, Ret_Val => #Ready5)
   END_RUNG
   // the same network as SCL:
   IF #At210 THEN
       #Ready5 := "F_PressDemoConfirmScrap"(SourcePath := #SourcePath, Seq := #Seq, AlarmLog := #AlarmLog);
   END_IF;
END_REGION

REGION Network 65
   RUNG wire#powerrail
      Contact( #At210 )
      "FRK_SeqReady"(Ok1 := #Ready5, Ok2 := TRUE, Ok3 := TRUE, Ok4 := TRUE, Ok5 := TRUE, Seq := #Seq)
   END_RUNG
   // the same network as SCL:
   IF #At210 THEN
       "FRK_SeqReady"(Ok1 := #Ready5, Ok2 := TRUE, Ok3 := TRUE, Ok4 := TRUE, Ok5 := TRUE, Seq := #Seq);
   END_IF;
END_REGION

REGION Network 66
   RUNG wire#powerrail
      Contact( #At210 )
      "FRK_SeqRoute"(OnAdvance := 215, OnJump1 := -1, Seq := #Seq)
   END_RUNG
   // the same network as SCL:
   IF #At210 THEN "FRK_SeqRoute"(OnAdvance := 215, OnJump1 := -1, Seq := #Seq); END_IF;
END_REGION

REGION Network 67
   RUNG wire#powerrail
      "FRK_SeqAt"(StepNo := 215, Seq := #Seq, Ret_Val => #At215)
   END_RUNG
   // the same network as SCL:
   #At215 := "FRK_SeqAt"(StepNo := 215, Seq := #Seq);
END_REGION

REGION Network 68
   RUNG wire#powerrail
      Contact( #At215 )
      "FRK_SeqStep"(StepNo := 215, StepName := 'project.step.pressScrapPart', Seq := #Seq, Row := #Row12)
   END_RUNG
   // the same network as SCL:
   IF #At215 THEN
       "FRK_SeqStep"(StepNo := 215, StepName := 'project.step.pressScrapPart', Seq := #Seq, Row := #Row12);
   END_IF;
END_REGION

REGION Network 69
   RUNG wire#powerrail
      Contact( #At215 )
      "F_PressDemoScrap"(Seq := #Seq, Cycle := #Cycle, Core := #Core, Unit := #Unit, Status := #Status, Part := #Part, AlarmLog := #AlarmLog, Ret_Val => #Ready5)
   END_RUNG
   // the same network as SCL:
   IF #At215 THEN
       #Ready5 := "F_PressDemoScrap"(Seq := #Seq,
                               Cycle := #Cycle,
                               Core := #Core,
                               Unit := #Unit,
                               Status := #Status,
                               Part := #Part,
                               AlarmLog := #AlarmLog);
   END_IF;
END_REGION

REGION Network 70
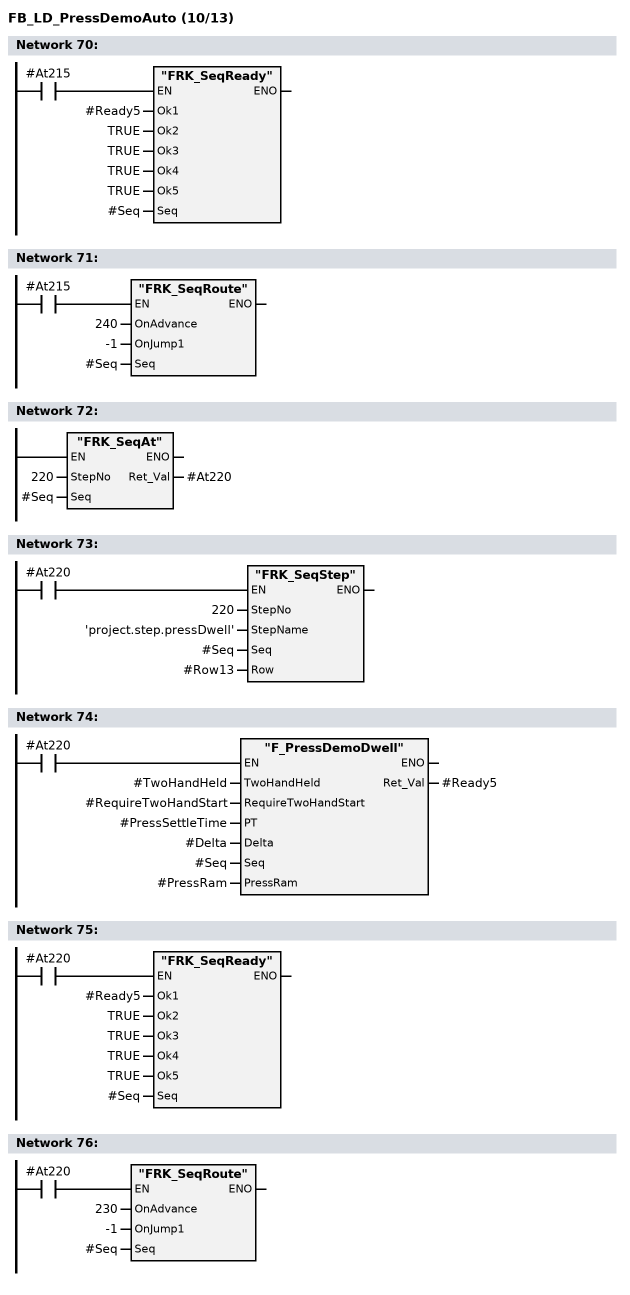
   RUNG wire#powerrail
      Contact( #At215 )
      "FRK_SeqReady"(Ok1 := #Ready5, Ok2 := TRUE, Ok3 := TRUE, Ok4 := TRUE, Ok5 := TRUE, Seq := #Seq)
   END_RUNG
   // the same network as SCL:
   IF #At215 THEN
       "FRK_SeqReady"(Ok1 := #Ready5, Ok2 := TRUE, Ok3 := TRUE, Ok4 := TRUE, Ok5 := TRUE, Seq := #Seq);
   END_IF;
END_REGION

REGION Network 71
   RUNG wire#powerrail
      Contact( #At215 )
      "FRK_SeqRoute"(OnAdvance := 240, OnJump1 := -1, Seq := #Seq)
   END_RUNG
   // the same network as SCL:
   IF #At215 THEN "FRK_SeqRoute"(OnAdvance := 240, OnJump1 := -1, Seq := #Seq); END_IF;
END_REGION

REGION Network 72
   RUNG wire#powerrail
      "FRK_SeqAt"(StepNo := 220, Seq := #Seq, Ret_Val => #At220)
   END_RUNG
   // the same network as SCL:
   #At220 := "FRK_SeqAt"(StepNo := 220, Seq := #Seq);
END_REGION

REGION Network 73
   RUNG wire#powerrail
      Contact( #At220 )
      "FRK_SeqStep"(StepNo := 220, StepName := 'project.step.pressDwell', Seq := #Seq, Row := #Row13)
   END_RUNG
   // the same network as SCL:
   IF #At220 THEN
       "FRK_SeqStep"(StepNo := 220, StepName := 'project.step.pressDwell', Seq := #Seq, Row := #Row13);
   END_IF;
END_REGION

REGION Network 74
   RUNG wire#powerrail
      Contact( #At220 )
      "F_PressDemoDwell"(TwoHandHeld := #TwoHandHeld, RequireTwoHandStart := #RequireTwoHandStart, PT := #PressSettleTime, Delta := #Delta, Seq := #Seq, PressRam := #PressRam, Ret_Val => #Ready5)
   END_RUNG
   // the same network as SCL:
   IF #At220 THEN
       #Ready5 := "F_PressDemoDwell"(TwoHandHeld := #TwoHandHeld,
                               RequireTwoHandStart := #RequireTwoHandStart,
                               PT := #PressSettleTime,
                               Delta := #Delta,
                               Seq := #Seq,
                               PressRam := #PressRam);
   END_IF;
END_REGION

REGION Network 75
   RUNG wire#powerrail
      Contact( #At220 )
      "FRK_SeqReady"(Ok1 := #Ready5, Ok2 := TRUE, Ok3 := TRUE, Ok4 := TRUE, Ok5 := TRUE, Seq := #Seq)
   END_RUNG
   // the same network as SCL:
   IF #At220 THEN
       "FRK_SeqReady"(Ok1 := #Ready5, Ok2 := TRUE, Ok3 := TRUE, Ok4 := TRUE, Ok5 := TRUE, Seq := #Seq);
   END_IF;
END_REGION

REGION Network 76
   RUNG wire#powerrail
      Contact( #At220 )
      "FRK_SeqRoute"(OnAdvance := 230, OnJump1 := -1, Seq := #Seq)
   END_RUNG
   // the same network as SCL:
   IF #At220 THEN "FRK_SeqRoute"(OnAdvance := 230, OnJump1 := -1, Seq := #Seq); END_IF;
END_REGION

REGION Network 77
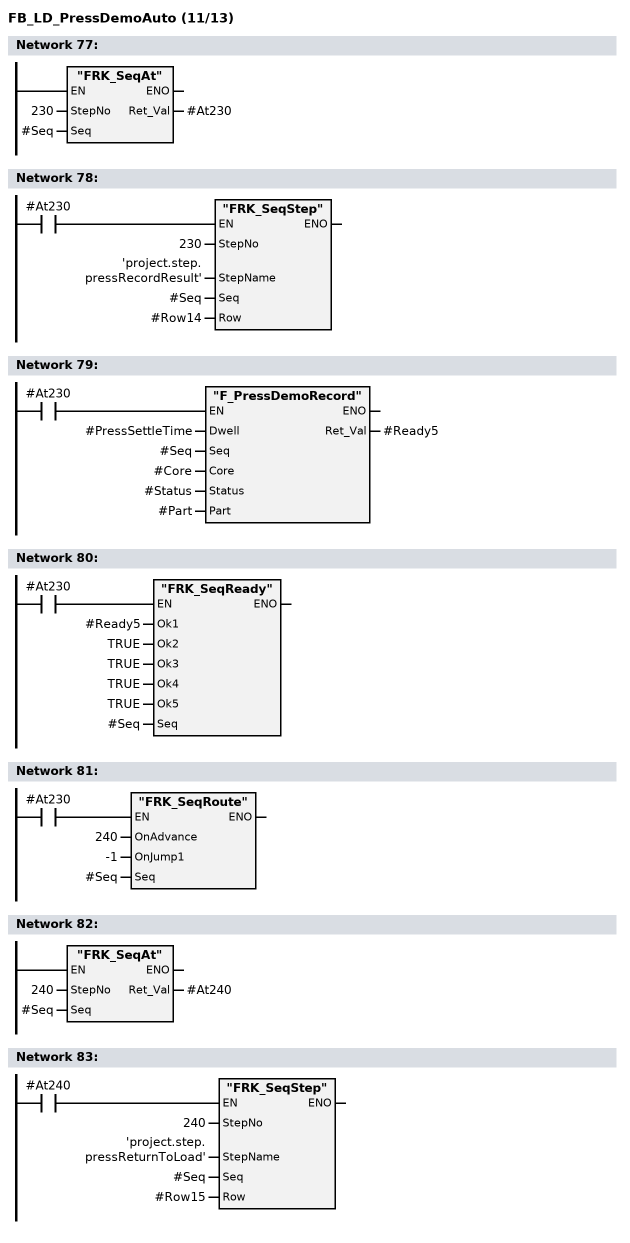
   RUNG wire#powerrail
      "FRK_SeqAt"(StepNo := 230, Seq := #Seq, Ret_Val => #At230)
   END_RUNG
   // the same network as SCL:
   #At230 := "FRK_SeqAt"(StepNo := 230, Seq := #Seq);
END_REGION

REGION Network 78
   RUNG wire#powerrail
      Contact( #At230 )
      "FRK_SeqStep"(StepNo := 230, StepName := 'project.step.pressRecordResult', Seq := #Seq, Row := #Row14)
   END_RUNG
   // the same network as SCL:
   IF #At230 THEN
       "FRK_SeqStep"(StepNo := 230, StepName := 'project.step.pressRecordResult', Seq := #Seq, Row := #Row14);
   END_IF;
END_REGION

REGION Network 79
   RUNG wire#powerrail
      Contact( #At230 )
      "F_PressDemoRecord"(Dwell := #PressSettleTime, Seq := #Seq, Core := #Core, Status := #Status, Part := #Part, Ret_Val => #Ready5)
   END_RUNG
   // the same network as SCL:
   IF #At230 THEN
       #Ready5 := "F_PressDemoRecord"(Dwell := #PressSettleTime,
                               Seq := #Seq,
                               Core := #Core,
                               Status := #Status,
                               Part := #Part);
   END_IF;
END_REGION

REGION Network 80
   RUNG wire#powerrail
      Contact( #At230 )
      "FRK_SeqReady"(Ok1 := #Ready5, Ok2 := TRUE, Ok3 := TRUE, Ok4 := TRUE, Ok5 := TRUE, Seq := #Seq)
   END_RUNG
   // the same network as SCL:
   IF #At230 THEN
       "FRK_SeqReady"(Ok1 := #Ready5, Ok2 := TRUE, Ok3 := TRUE, Ok4 := TRUE, Ok5 := TRUE, Seq := #Seq);
   END_IF;
END_REGION

REGION Network 81
   RUNG wire#powerrail
      Contact( #At230 )
      "FRK_SeqRoute"(OnAdvance := 240, OnJump1 := -1, Seq := #Seq)
   END_RUNG
   // the same network as SCL:
   IF #At230 THEN "FRK_SeqRoute"(OnAdvance := 240, OnJump1 := -1, Seq := #Seq); END_IF;
END_REGION

REGION Network 82
   RUNG wire#powerrail
      "FRK_SeqAt"(StepNo := 240, Seq := #Seq, Ret_Val => #At240)
   END_RUNG
   // the same network as SCL:
   #At240 := "FRK_SeqAt"(StepNo := 240, Seq := #Seq);
END_REGION

REGION Network 83
   RUNG wire#powerrail
      Contact( #At240 )
      "FRK_SeqStep"(StepNo := 240, StepName := 'project.step.pressReturnToLoad', Seq := #Seq, Row := #Row15)
   END_RUNG
   // the same network as SCL:
   IF #At240 THEN
       "FRK_SeqStep"(StepNo := 240, StepName := 'project.step.pressReturnToLoad', Seq := #Seq, Row := #Row15);
   END_IF;
END_REGION

REGION Network 84
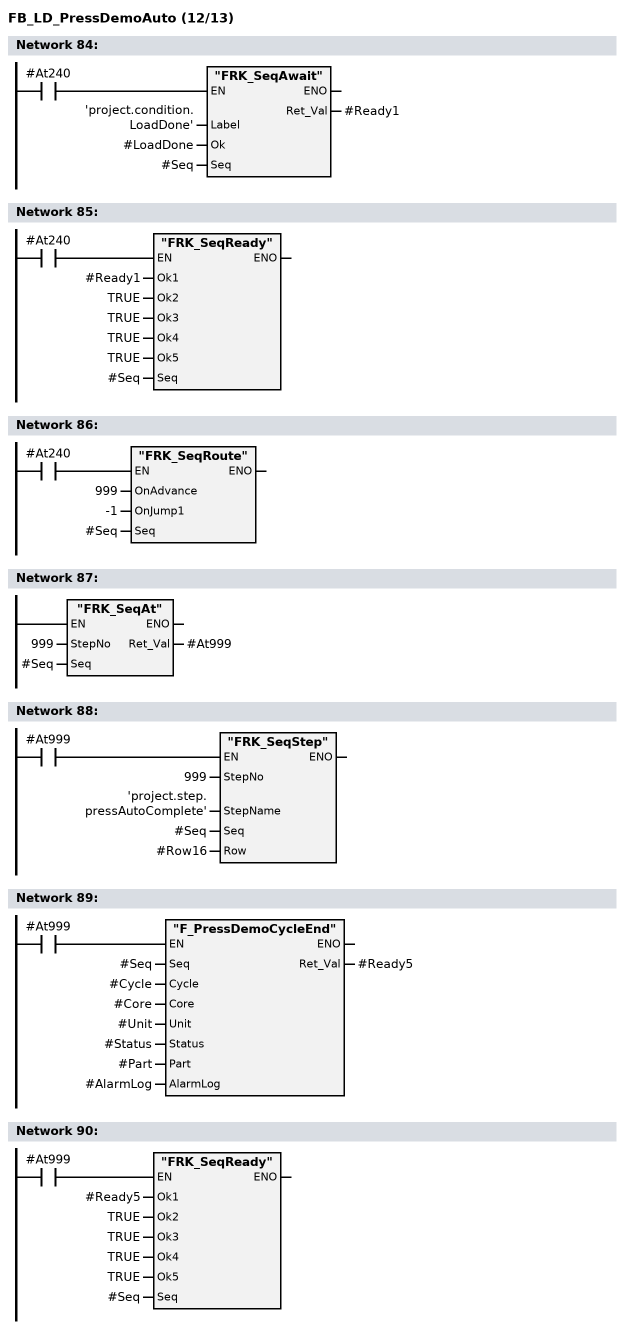
   RUNG wire#powerrail
      Contact( #At240 )
      "FRK_SeqAwait"(Label := 'project.condition.LoadDone', Ok := #LoadDone, Seq := #Seq, Ret_Val => #Ready1)
   END_RUNG
   // the same network as SCL:
   IF #At240 THEN
       #Ready1 := "FRK_SeqAwait"(Label := 'project.condition.LoadDone', Ok := #LoadDone, Seq := #Seq);
   END_IF;
END_REGION

REGION Network 85
   RUNG wire#powerrail
      Contact( #At240 )
      "FRK_SeqReady"(Ok1 := #Ready1, Ok2 := TRUE, Ok3 := TRUE, Ok4 := TRUE, Ok5 := TRUE, Seq := #Seq)
   END_RUNG
   // the same network as SCL:
   IF #At240 THEN
       "FRK_SeqReady"(Ok1 := #Ready1, Ok2 := TRUE, Ok3 := TRUE, Ok4 := TRUE, Ok5 := TRUE, Seq := #Seq);
   END_IF;
END_REGION

REGION Network 86
   RUNG wire#powerrail
      Contact( #At240 )
      "FRK_SeqRoute"(OnAdvance := 999, OnJump1 := -1, Seq := #Seq)
   END_RUNG
   // the same network as SCL:
   IF #At240 THEN "FRK_SeqRoute"(OnAdvance := 999, OnJump1 := -1, Seq := #Seq); END_IF;
END_REGION

REGION Network 87
   RUNG wire#powerrail
      "FRK_SeqAt"(StepNo := 999, Seq := #Seq, Ret_Val => #At999)
   END_RUNG
   // the same network as SCL:
   #At999 := "FRK_SeqAt"(StepNo := 999, Seq := #Seq);
END_REGION

REGION Network 88
   RUNG wire#powerrail
      Contact( #At999 )
      "FRK_SeqStep"(StepNo := 999, StepName := 'project.step.pressAutoComplete', Seq := #Seq, Row := #Row16)
   END_RUNG
   // the same network as SCL:
   IF #At999 THEN
       "FRK_SeqStep"(StepNo := 999, StepName := 'project.step.pressAutoComplete', Seq := #Seq, Row := #Row16);
   END_IF;
END_REGION

REGION Network 89
   RUNG wire#powerrail
      Contact( #At999 )
      "F_PressDemoCycleEnd"(Seq := #Seq, Cycle := #Cycle, Core := #Core, Unit := #Unit, Status := #Status, Part := #Part, AlarmLog := #AlarmLog, Ret_Val => #Ready5)
   END_RUNG
   // the same network as SCL:
   IF #At999 THEN
       #Ready5 := "F_PressDemoCycleEnd"(Seq := #Seq,
                               Cycle := #Cycle,
                               Core := #Core,
                               Unit := #Unit,
                               Status := #Status,
                               Part := #Part,
                               AlarmLog := #AlarmLog);
   END_IF;
END_REGION

REGION Network 90
   RUNG wire#powerrail
      Contact( #At999 )
      "FRK_SeqReady"(Ok1 := #Ready5, Ok2 := TRUE, Ok3 := TRUE, Ok4 := TRUE, Ok5 := TRUE, Seq := #Seq)
   END_RUNG
   // the same network as SCL:
   IF #At999 THEN
       "FRK_SeqReady"(Ok1 := #Ready5, Ok2 := TRUE, Ok3 := TRUE, Ok4 := TRUE, Ok5 := TRUE, Seq := #Seq);
   END_IF;
END_REGION

REGION Network 91
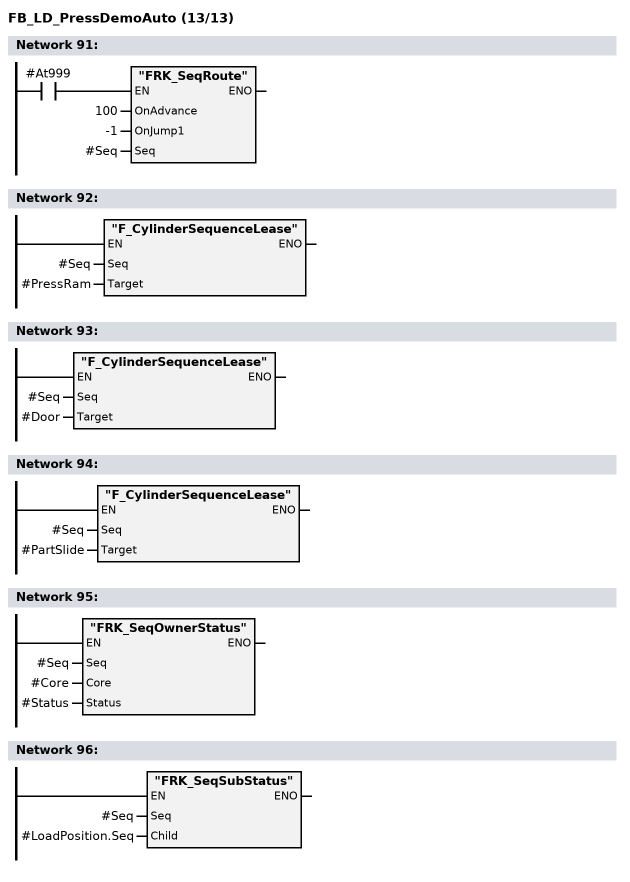
   RUNG wire#powerrail
      Contact( #At999 )
      "FRK_SeqRoute"(OnAdvance := 100, OnJump1 := -1, Seq := #Seq)
   END_RUNG
   // the same network as SCL:
   IF #At999 THEN "FRK_SeqRoute"(OnAdvance := 100, OnJump1 := -1, Seq := #Seq); END_IF;
END_REGION

REGION Network 92
   RUNG wire#powerrail
      "F_CylinderSequenceLease"(Seq := #Seq, Target := #PressRam)
   END_RUNG
   // the same network as SCL:
   "F_CylinderSequenceLease"(Seq := #Seq, Target := #PressRam);
END_REGION

REGION Network 93
   RUNG wire#powerrail
      "F_CylinderSequenceLease"(Seq := #Seq, Target := #Door)
   END_RUNG
   // the same network as SCL:
   "F_CylinderSequenceLease"(Seq := #Seq, Target := #Door);
END_REGION

REGION Network 94
   RUNG wire#powerrail
      "F_CylinderSequenceLease"(Seq := #Seq, Target := #PartSlide)
   END_RUNG
   // the same network as SCL:
   "F_CylinderSequenceLease"(Seq := #Seq, Target := #PartSlide);
END_REGION

REGION Network 95
   RUNG wire#powerrail
      "FRK_SeqOwnerStatus"(Seq := #Seq, Core := #Core, Status := #Status)
   END_RUNG
   // the same network as SCL:
   "FRK_SeqOwnerStatus"(Seq := #Seq, Core := #Core, Status := #Status);
END_REGION

REGION Network 96
   RUNG wire#powerrail
      "FRK_SeqSubStatus"(Seq := #Seq, Child := #LoadPosition.Seq)
   END_RUNG
   // the same network as SCL:
   "FRK_SeqSubStatus"(Seq := #Seq, Child := #LoadPosition.Seq);
END_REGION
END_FUNCTION_BLOCK

FUNCTION "FRK_SeqBegin" : Void   // FC124, SCL
{ S7_Optimized_Access := 'TRUE' }
VERSION : 0.1
// Shared sequence services. The examples generator binds Core enum constants.
// stored: AutoNumber true, IsIECCheckEnabled false, SetENOAutomatically false, UDAEnableTagReadback false
   VAR_INPUT
      Run : Bool;
      Reset : Bool;
      OwnerIndex : DInt;
      ChainIndex : DInt;
      BranchIndex : DInt;
      Delta : Time;
   END_VAR
   VAR_IN_OUT
      Seq : "FRK_SequenceCtx";
   END_VAR
BEGIN

   #Seq.Scan := #Seq.Scan + 1;
   #Seq.Restart := #Reset OR (#Run AND NOT #Seq.RunPrevious);
   #Seq.RunPrevious := #Run;
   #Seq.OwnerIndex := #OwnerIndex;
   #Seq.ChainIndex := #ChainIndex;
   #Seq.BranchIndex := #BranchIndex;
   #Seq.RetVal := 0;
   #Seq.Pending := FALSE;
   #Seq.CommandFailed := FALSE;
   #Seq.CommandIssued := FALSE;
   #Seq.Awaiting := '';
   IF NOT #Run OR #Seq.Restart THEN
       #Seq.Step := 0;
       #Seq.RecordedStep := -1;
       #Seq.Visit := #Seq.Visit + 1;
       #Seq.Done := FALSE;
       #Seq.Error := FALSE;
       #Seq.StartLatched := FALSE;
       #Seq.Elapsed := T#0ms;
       #Seq.DelayElapsed := T#0ms;
       #Seq.ErrorDiagnostic.ReasonCode := 0;
   END_IF;
   #Seq.Running := #Run AND NOT #Seq.Done AND NOT #Seq.Error
   AND #OwnerIndex > 0 AND #ChainIndex > 0;
   #Seq.ScanStep := #Seq.Step;
   IF #Seq.Running AND #Delta > T#0ms THEN
       #Seq.Elapsed := #Seq.Elapsed + #Delta;
   END_IF;
END_FUNCTION

FUNCTION "FRK_SeqStart" : Void   // FC125, SCL
{ S7_Optimized_Access := 'TRUE' }
VERSION : 0.1
// stored: AutoNumber true, IsIECCheckEnabled false, SetENOAutomatically false, UDAEnableTagReadback false
   VAR_INPUT
      StartPulse : Bool;
   END_VAR
   VAR_IN_OUT
      Seq : "FRK_SequenceCtx";
   END_VAR
BEGIN

   IF #Seq.Running THEN
       #Seq.StartLatched := #Seq.StartLatched OR #StartPulse;
   END_IF;
END_FUNCTION

FUNCTION "F_PressDemoReset" : Void   // FC159, SCL
{ S7_Optimized_Access := 'TRUE' }
VERSION : 0.1
// Project policy only. Lifecycle, ownership, waits, messages and once-per-visit
//  bookkeeping stay in Core; GRAPH actions and the ST/LD twins call these FCs.
// stored: AutoNumber true, IsIECCheckEnabled false, SetENOAutomatically false, UDAEnableTagReadback false
   VAR_IN_OUT
      Seq : "FRK_SequenceCtx";
      Cycle : "ST_PressDemoCycle";
   END_VAR
BEGIN

   IF #Seq.Restart THEN
       #Cycle.PartInMachine := FALSE;
       #Cycle.PartDispositioned := FALSE;
       #Cycle.CycleCompleted := FALSE;
       #Cycle.FailureReason := 0;
   END_IF;
END_FUNCTION

FUNCTION "FRK_SeqSubActive" : Bool   // FC136, SCL
{ S7_Optimized_Access := 'TRUE' }
VERSION : 0.1
// stored: AutoNumber true, IsIECCheckEnabled false, SetENOAutomatically false, UDAEnableTagReadback false
   VAR_INPUT
      Run : Bool;
      StepNo : DInt;
   END_VAR
   VAR_IN_OUT
      Seq : "FRK_SequenceCtx";
   END_VAR
BEGIN

   #FRK_SeqSubActive := #Run AND #Seq.Running AND NOT #Seq.Error AND #Seq.Step = #StepNo;
END_FUNCTION

FUNCTION "F_PressDemoLoadPosition" : Bool   // FC170, SCL
{ S7_Optimized_Access := 'TRUE' }
VERSION : 0.1
// stored: AutoNumber true, IsIECCheckEnabled false, SetENOAutomatically false, UDAEnableTagReadback false
   VAR_INPUT
      Run : Bool;
      Reset : Bool;
      OwnerIndex : DInt;
      Delta : Time;
   END_VAR
   VAR_IN_OUT
      Target : "FB_PressDemoLoadPosition";
      PressRam : "FB_CylinderCM";
      Door : "FB_CylinderCM";
      PartSlide : "FB_CylinderCM";
   END_VAR
BEGIN

   #Target(Run := #Run,
           Reset := #Reset,
           OwnerIndex := #OwnerIndex,
           Delta := #Delta,
           PressRam := #PressRam,
           Door := #Door,
           PartSlide := #PartSlide);
   #F_PressDemoLoadPosition := #Target.Seq.Done;
END_FUNCTION

FUNCTION "F_CylinderSequenceLease" : Void   // FC156, SCL
{ S7_Optimized_Access := 'TRUE' }
VERSION : 0.1
// stored: AutoNumber true, IsIECCheckEnabled false, SetENOAutomatically false, UDAEnableTagReadback false
   VAR_IN_OUT
      Seq : "FRK_SequenceCtx";
      Target : "FB_CylinderCM";
   END_VAR
BEGIN

   IF #Target.Device.Lease.OwnerIndex = #Seq.OwnerIndex
       AND #Target.Device.Lease.ChainIndex = #Seq.ChainIndex
       AND #Target.Device.Lease.BranchIndex = #Seq.BranchIndex
       AND #Seq.OwnerIndex > 0 AND #Seq.ChainIndex > 0
       AND (NOT #Seq.Running OR #Seq.Error OR #Seq.Restart) THEN
       #Target.Device.Withdrawn := TRUE;
   END_IF;
   IF #Target.Device.Lease.OwnerIndex = #Seq.OwnerIndex
       AND #Target.Device.Lease.ChainIndex = #Seq.ChainIndex
       AND #Target.Device.Lease.BranchIndex = #Seq.BranchIndex
       AND #Target.Device.Lease.AbortIssued AND #Target.Device.Lease.ReleasedScan <> #Seq.Scan THEN
       #Target.Abort := FALSE;
       #Target.Device.Lease.AbortIssued := FALSE;
   END_IF;
   IF #Target.Device.Lease.Raised AND #Target.Device.Lease.OwnerIndex = #Seq.OwnerIndex
       AND #Target.Device.Lease.ChainIndex = #Seq.ChainIndex
       AND #Target.Device.Lease.BranchIndex = #Seq.BranchIndex
       AND (NOT #Seq.Running OR #Seq.Error OR #Seq.Restart OR #Target.Device.Lease.Step <> #Seq.Step) THEN
       #Target.Abort := #Target.Busy;
       #Target.Device.Lease.AbortIssued := #Target.Busy;
   END_IF;
   "FRK_SeqLease"(Seq := #Seq,
                  Lease := #Target.Device.Lease,
                  Execute := #Target.Execute);
END_FUNCTION

FUNCTION "FRK_SeqOwnerStatus" : Void   // FC141, SCL
{ S7_Optimized_Access := 'TRUE' }
VERSION : 0.1
// stored: AutoNumber true, IsIECCheckEnabled false, SetENOAutomatically false, UDAEnableTagReadback false
   VAR_IN_OUT
      Seq : "FRK_SequenceCtx";
      Core : "FRK_Core";
      Status : "ST_ModuleStatus";
   END_VAR
BEGIN

   IF #Core.Exec = 3 THEN
       #Seq.Error := TRUE;
       #Seq.ErrorDiagnostic := #Status.Diagnostic;
   ELSIF #Seq.Error THEN
       "FRK_AdoptFault"(Core := #Core,
                        Status := #Status,
                        Diag := #Seq.ErrorDiagnostic);
   END_IF;
END_FUNCTION

FUNCTION "FRK_SeqSubStatus" : Void   // FC137, SCL
{ S7_Optimized_Access := 'TRUE' }
VERSION : 0.1
// stored: AutoNumber true, IsIECCheckEnabled false, SetENOAutomatically false, UDAEnableTagReadback false
   VAR_IN_OUT
      Seq : "FRK_SequenceCtx";
      Child : "FRK_SequenceCtx";
   END_VAR
BEGIN

   IF #Child.Error THEN
       #Seq.Error := TRUE;
       #Seq.ErrorDiagnostic := #Child.ErrorDiagnostic;
   END_IF;
END_FUNCTION

FUNCTION "FRK_SeqAt" : Bool   // FC128, SCL
{ S7_Optimized_Access := 'TRUE' }
VERSION : 0.1
// stored: AutoNumber true, IsIECCheckEnabled false, SetENOAutomatically false, UDAEnableTagReadback false
   VAR_INPUT
      StepNo : DInt;
   END_VAR
   VAR_IN_OUT
      Seq : "FRK_SequenceCtx";
   END_VAR
BEGIN

   // Capture dispatch once: a forward LD transition cannot execute the next
   // state's rung in this scan or hide an Execute-low reset scan.
   #FRK_SeqAt := #Seq.Running AND NOT #Seq.Error AND #Seq.ScanStep = #StepNo;
END_FUNCTION

FUNCTION "FRK_SeqStep" : Void   // FC129, SCL
{ S7_Optimized_Access := 'TRUE' }
VERSION : 0.1
// stored: AutoNumber true, IsIECCheckEnabled false, SetENOAutomatically false, UDAEnableTagReadback false
   VAR_INPUT
      StepNo : DInt;
      StepName : String;
   END_VAR
   VAR_IN_OUT
      Seq : "FRK_SequenceCtx";
      Row : "FRK_SequenceRow";
   END_VAR
BEGIN

   IF #Seq.RecordedStep <> #StepNo THEN
       #Seq.Visit := #Seq.Visit + 1;
       #Seq.Elapsed := T#0ms;
       #Seq.DelayElapsed := T#0ms;
       #Seq.RecordedStep := #StepNo;
       #Seq.Warned := FALSE;
   END_IF;
   #Seq.Step := #StepNo;
   #Seq.StepName := #StepName;
   #Row.StepNo := #StepNo;
   #Row.Visited := TRUE;
   #Row.LastDuration := #Seq.Elapsed;
END_FUNCTION

FUNCTION "FRK_SeqReady" : Void   // FC138, SCL
{ S7_Optimized_Access := 'TRUE' }
VERSION : 0.1
// stored: AutoNumber true, IsIECCheckEnabled false, SetENOAutomatically false, UDAEnableTagReadback false
   VAR_INPUT
      Ok1 : Bool;
      Ok2 : Bool;
      Ok3 : Bool;
      Ok4 : Bool;
      Ok5 : Bool;
   END_VAR
   VAR_IN_OUT
      Seq : "FRK_SequenceCtx";
   END_VAR
BEGIN

   "FRK_SeqSelect"(Seq := #Seq, AdvanceOk := #Ok1 AND #Ok2 AND #Ok3 AND #Ok4 AND #Ok5, Jump1Ok := FALSE);
END_FUNCTION

FUNCTION "FRK_SeqRoute" : Void   // FC142, SCL
{ S7_Optimized_Access := 'TRUE' }
VERSION : 0.1
// stored: AutoNumber true, IsIECCheckEnabled false, SetENOAutomatically false, UDAEnableTagReadback false
   VAR_INPUT
      OnAdvance : DInt;
      OnJump1 : DInt;
   END_VAR
   VAR_IN_OUT
      Seq : "FRK_SequenceCtx";
   END_VAR
BEGIN

   IF NOT #Seq.Running OR #Seq.Error THEN
       RETURN;
   END_IF;
   CASE #Seq.RetVal OF
       1:
           IF #OnAdvance >= 0 THEN
               #Seq.Step := #OnAdvance;
           END_IF;
       2:
           IF #OnJump1 >= 0 THEN
               #Seq.Step := #OnJump1;
           END_IF;
       ELSE
           RETURN;
   END_CASE;
END_FUNCTION

FUNCTION "F_PressDemoAwaitCycle" : Bool   // FC160, SCL
{ S7_Optimized_Access := 'TRUE' }
VERSION : 0.1
// stored: AutoNumber true, IsIECCheckEnabled false, SetENOAutomatically false, UDAEnableTagReadback false
   VAR_INPUT
      PartPresent : Bool;
      PartQuality : Bool;
      AirPressureOk : Bool;
      RequireTwoHandStart : Bool;
   END_VAR
   VAR_IN_OUT
      Seq : "FRK_SequenceCtx";
      Cycle : "ST_PressDemoCycle";
      Core : "FRK_Core";
      Unit : "FRK_Unit";
      Status : "ST_ModuleStatus";
      Part : "ST_PartContext";
      AlarmLog : "FRK_AlarmLog";
   END_VAR
   VAR_TEMP
      PartReady : Bool;
      AirReady : Bool;
      StartReady : Bool;
      Received : Bool;
   END_VAR
BEGIN

   #F_PressDemoAwaitCycle := FALSE;
   #Cycle.CycleCompleted := FALSE;
   IF #Unit.StopReq THEN
       "FRK_Complete"(Core := #Core,
                      Status := #Status);
       "FRK_SeqComplete"(Seq := #Seq);
       RETURN;
   END_IF;
   #PartReady := "FRK_SeqAwait"(Seq := #Seq, Label := 'project.condition.partPresent', Ok := #PartPresent AND #PartQuality);
   #AirReady := "FRK_SeqAwait"(Seq := #Seq, Label := 'project.condition.airPressureOk', Ok := #AirPressureOk);
   #StartReady := "FRK_SeqAwait"(Seq := #Seq, Label := 'project.condition.twoHandStart', Ok := #Seq.StartLatched OR NOT #RequireTwoHandStart);
   IF NOT (#PartReady AND #AirReady AND #StartReady) THEN
       RETURN;
   END_IF;
   IF NOT #Cycle.PartInMachine THEN
       #Received := "FRK_PartReceived"(Core := #Core, Unit := #Unit, Status := #Status, Part := #Part, AlarmLog := #AlarmLog);
       IF #Core.Exec = 3 THEN
           #Seq.Error := TRUE;
           #Seq.ErrorDiagnostic := #Status.Diagnostic;
           RETURN;
       END_IF;
       #Cycle.PartInMachine := TRUE;
   END_IF;
   #F_PressDemoAwaitCycle := TRUE;
END_FUNCTION

FUNCTION "F_CylinderRetract" : Bool   // FC155, SCL
{ S7_Optimized_Access := 'TRUE' }
VERSION : 0.1
// stored: AutoNumber true, IsIECCheckEnabled false, SetENOAutomatically false, UDAEnableTagReadback false
   VAR_IN_OUT
      Seq : "FRK_SequenceCtx";
      Target : "FB_CylinderCM";
   END_VAR
BEGIN

   #F_CylinderRetract := "FRK_SeqCommand"(Seq := #Seq, Lease := #Target.Device.Lease,
                                          Execute := #Target.Execute, Command := #Target.Command,
                                          Value := 2, Label := 'Cylinder.RETRACT', Ready := #Target.Status.State = 0,
                                          Done := #Target.Done, Error := #Target.Error, OwnFailure := FALSE, Diagnostic := #Target.Status.Diagnostic);
END_FUNCTION

FUNCTION "F_CylinderExtend" : Bool   // FC153, SCL
{ S7_Optimized_Access := 'TRUE' }
VERSION : 0.1
// The typed device API owns handshake access; sequence authors call actions.
// stored: AutoNumber true, IsIECCheckEnabled false, SetENOAutomatically false, UDAEnableTagReadback false
   VAR_IN_OUT
      Seq : "FRK_SequenceCtx";
      Target : "FB_CylinderCM";
   END_VAR
BEGIN

   #F_CylinderExtend := "FRK_SeqCommand"(Seq := #Seq, Lease := #Target.Device.Lease,
                                         Execute := #Target.Execute, Command := #Target.Command,
                                         Value := 1, Label := 'Cylinder.EXTEND', Ready := #Target.Status.State = 0,
                                         Done := #Target.Done, Error := #Target.Error, OwnFailure := FALSE, Diagnostic := #Target.Status.Diagnostic);
END_FUNCTION

FUNCTION "F_PressDemoStarted" : Void   // FC161, SCL
{ S7_Optimized_Access := 'TRUE' }
VERSION : 0.1
// stored: AutoNumber true, IsIECCheckEnabled false, SetENOAutomatically false, UDAEnableTagReadback false
   VAR_IN_OUT
      Seq : "FRK_SequenceCtx";
      Unit : "FRK_Unit";
      Status : "ST_ModuleStatus";
      Part : "ST_PartContext";
      AlarmLog : "FRK_AlarmLog";
   END_VAR
BEGIN

   IF "FRK_SeqOnce"(Seq := #Seq, Enable := #Seq.CommandIssued, Token := #Seq.Step) THEN
       "FRK_PartStarted"(Unit := #Unit,
                         Status := #Status,
                         Part := #Part,
                         AlarmLog := #AlarmLog);
   END_IF;
END_FUNCTION

FUNCTION "FRK_SeqDelay" : Bool   // FC131, SCL
{ S7_Optimized_Access := 'TRUE' }
VERSION : 0.1
// stored: AutoNumber true, IsIECCheckEnabled false, SetENOAutomatically false, UDAEnableTagReadback false
   VAR_INPUT
      Permit : Bool;
      PT : Time;
      Delta : Time;
   END_VAR
   VAR_IN_OUT
      Seq : "FRK_SequenceCtx";
   END_VAR
BEGIN

   IF #Permit AND #Delta > T#0ms THEN
       #Seq.DelayElapsed := #Seq.DelayElapsed + #Delta;
   END_IF;
   #FRK_SeqDelay := #Permit AND #Seq.DelayElapsed >= #PT;
END_FUNCTION

FUNCTION "F_PressDemoDoorClose" : Void   // FC162, SCL
{ S7_Optimized_Access := 'TRUE' }
VERSION : 0.1
// stored: AutoNumber true, IsIECCheckEnabled false, SetENOAutomatically false, UDAEnableTagReadback false
   VAR_INPUT
      Closed : Bool;
      TwoHandHeld : Bool;
      RequireTwoHandStart : Bool;
      SourcePath : String;
   END_VAR
   VAR_IN_OUT
      Seq : "FRK_SequenceCtx";
      AlarmLog : "FRK_AlarmLog";
   END_VAR
   VAR_TEMP
      Held : Bool;
      Diag : "ST_Diagnostic";
   END_VAR
BEGIN

   #Held := "FRK_SeqAwait"(Seq := #Seq, Label := 'project.condition.twoHandHeldDuringDoorClose', Ok := #TwoHandHeld OR NOT #RequireTwoHandStart);
   "FRK_SeqSelect"(Seq := #Seq,
                   AdvanceOk := #Closed,
                   Jump1Ok := NOT #Held);
   IF #Seq.RetVal = 2 THEN
       #Diag := "FRK_UnitScratch".EmptyDiagnostic;
       #Diag.ReasonCode := 12001;
       #Diag.Description := WSTRING#'project.warning.twoHandReleasedDuringDoorClose';
       #Diag.SourcePath := STRING_TO_WSTRING(#SourcePath);
       #Diag.Severity := 0;
       #Diag.Category := 0;
       "FRK_SeqMessage"(Seq := #Seq,
                        AlarmLog := #AlarmLog,
                        Diag := #Diag);
   END_IF;
END_FUNCTION

FUNCTION "F_PressDemoClearStart" : Void   // FC163, SCL
{ S7_Optimized_Access := 'TRUE' }
VERSION : 0.1
// stored: AutoNumber true, IsIECCheckEnabled false, SetENOAutomatically false, UDAEnableTagReadback false
   VAR_INPUT
      Complete : Bool;
   END_VAR
   VAR_IN_OUT
      Seq : "FRK_SequenceCtx";
   END_VAR
BEGIN

   IF #Complete THEN
       "FRK_SeqCycleEnd"(Seq := #Seq);
   END_IF;
END_FUNCTION

FUNCTION "F_CylinderExtendHandled" : Bool   // FC154, SCL
{ S7_Optimized_Access := 'TRUE' }
VERSION : 0.1
// The step deliberately owns a failure branch. The shared command service
//  still verifies ownership; the original child first-out is retained verbatim.
// stored: AutoNumber true, IsIECCheckEnabled false, SetENOAutomatically false, UDAEnableTagReadback false
   VAR_IN_OUT
      Seq : "FRK_SequenceCtx";
      Target : "FB_CylinderCM";
   END_VAR
BEGIN

   #F_CylinderExtendHandled := "FRK_SeqCommand"(Seq := #Seq, Lease := #Target.Device.Lease,
                                                Execute := #Target.Execute, Command := #Target.Command, Value := 1,
                                                Label := 'Cylinder.EXTEND', Ready := #Target.Status.State = 0,
                                                Done := #Target.Done, Error := #Target.Error, OwnFailure := TRUE, Diagnostic := #Target.Status.Diagnostic);
   "FRK_SeqHandled"(Seq := #Seq,
                    ChildCore := #Target.Core);
   IF #Seq.CommandFailed THEN
       // Releasing the terminal handshake must not re-energize the failed
       // direction while the owning step awaits an operator decision.
       "F_CylinderForcePermit"(Target := #Target,
                               Permit := FALSE);
   END_IF;
END_FUNCTION

FUNCTION "F_PressDemoRamResult" : Void   // FC164, SCL
{ S7_Optimized_Access := 'TRUE' }
VERSION : 0.1
// stored: AutoNumber true, IsIECCheckEnabled false, SetENOAutomatically false, UDAEnableTagReadback false
   VAR_INPUT
      Reached : Bool;
   END_VAR
   VAR_IN_OUT
      Seq : "FRK_SequenceCtx";
      Cycle : "ST_PressDemoCycle";
      AlarmLog : "FRK_AlarmLog";
   END_VAR
BEGIN

   "FRK_SeqSelect"(Seq := #Seq,
                   AdvanceOk := #Reached,
                   Jump1Ok := #Seq.CommandFailed);
   IF #Seq.RetVal = 2 THEN
       #Cycle.FailureReason := #Seq.HandledDiagnostic.ReasonCode;
       "FRK_SeqMessage"(Seq := #Seq,
                        AlarmLog := #AlarmLog,
                        Diag := #Seq.HandledDiagnostic);
   END_IF;
END_FUNCTION

FUNCTION "F_PressDemoConfirmScrap" : Bool   // FC165, SCL
{ S7_Optimized_Access := 'TRUE' }
VERSION : 0.1
// stored: AutoNumber true, IsIECCheckEnabled false, SetENOAutomatically false, UDAEnableTagReadback false
   VAR_INPUT
      SourcePath : String;
   END_VAR
   VAR_IN_OUT
      Seq : "FRK_SequenceCtx";
      AlarmLog : "FRK_AlarmLog";
   END_VAR
   VAR_TEMP
      Request : "ST_DecisionRequest";
      Asked : Bool;
      Answer : Int;
      Ready : Bool;
   END_VAR
BEGIN

   #Request := "FRK_Decisions".EmptyRequest;
   #Request.Prompt := WSTRING#'project.decision.pressNotReached';
   #Request.Options[1] := 'project.decision.confirmScrapAndReturn';
   // Scrap is deliberate: no timeout and no default answer.
   #Asked := "FRK_DecisionAsk"(Owner := #Seq.OwnerIndex, OwnerPath := STRING_TO_WSTRING(#SourcePath), Request := #Request, AlarmLog := #AlarmLog);
   #Answer := 0;
   IF #Asked THEN
       #Answer := "FRK_DecisionTake"(Owner := #Seq.OwnerIndex, AlarmLog := #AlarmLog);
   END_IF;
   #Ready := "FRK_SeqAwait"(Seq := #Seq, Label := 'project.condition.pressFailureConfirmation', Ok := #Asked AND #Answer = 1);
   #F_PressDemoConfirmScrap := #Ready;
END_FUNCTION

FUNCTION "F_PressDemoScrap" : Bool   // FC166, SCL
{ S7_Optimized_Access := 'TRUE' }
VERSION : 0.1
// stored: AutoNumber true, IsIECCheckEnabled false, SetENOAutomatically false, UDAEnableTagReadback false
   VAR_IN_OUT
      Seq : "FRK_SequenceCtx";
      Cycle : "ST_PressDemoCycle";
      Core : "FRK_Core";
      Unit : "FRK_Unit";
      Status : "ST_ModuleStatus";
      Part : "ST_PartContext";
      AlarmLog : "FRK_AlarmLog";
   END_VAR
   VAR_TEMP
      Written : Bool;
   END_VAR
BEGIN

   IF "FRK_SeqOnce"(Seq := #Seq, Enable := TRUE, Token := #Seq.Step) THEN
       #Written := "FRK_PartProcessed"(Core := #Core, Unit := #Unit, Status := #Status, Part := #Part, AlarmLog := #AlarmLog,
                                       Verdict := 2, Reason := #Cycle.FailureReason);
       IF NOT #Written AND #Unit.CarrierIndex = 0 AND #Unit.Nok < UDINT#4294967295 THEN
           #Unit.Nok := #Unit.Nok + 1;
           #Unit.NokReason := #Cycle.FailureReason;
       END_IF;
       #Cycle.PartDispositioned := TRUE;
       #Cycle.PartInMachine := FALSE;
       #Cycle.CycleCompleted := FALSE;
   END_IF;
   #F_PressDemoScrap := #Core.Exec <> 3;
END_FUNCTION

FUNCTION "F_PressDemoDwell" : Bool   // FC167, SCL
{ S7_Optimized_Access := 'TRUE' }
VERSION : 0.1
// stored: AutoNumber true, IsIECCheckEnabled false, SetENOAutomatically false, UDAEnableTagReadback false
   VAR_INPUT
      TwoHandHeld : Bool;
      RequireTwoHandStart : Bool;
      PT : Time;
      Delta : Time;
   END_VAR
   VAR_IN_OUT
      Seq : "FRK_SequenceCtx";
      PressRam : "FB_CylinderCM";
   END_VAR
   VAR_TEMP
      Held : Bool;
   END_VAR
BEGIN

   #Held := "FRK_SeqAwait"(Seq := #Seq, Label := 'project.condition.twoHandHeldDuringPress', Ok := #TwoHandHeld OR NOT #RequireTwoHandStart);
   "F_CylinderForcePermit"(Target := #PressRam,
                           Permit := #Held);
   #F_PressDemoDwell := "FRK_SeqDelay"(Seq := #Seq, Permit := #Held, PT := #PT, Delta := #Delta);
END_FUNCTION

FUNCTION "F_PressDemoRecord" : Bool   // FC168, SCL
{ S7_Optimized_Access := 'TRUE' }
VERSION : 0.1
// stored: AutoNumber true, IsIECCheckEnabled false, SetENOAutomatically false, UDAEnableTagReadback false
   VAR_INPUT
      Dwell : Time;
   END_VAR
   VAR_IN_OUT
      Seq : "FRK_SequenceCtx";
      Core : "FRK_Core";
      Status : "ST_ModuleStatus";
      Part : "ST_PartContext";
   END_VAR
   VAR_TEMP
      Recorded : Bool;
   END_VAR
BEGIN

   IF "FRK_SeqOnce"(Seq := #Seq, Enable := TRUE, Token := #Seq.Step) THEN
       #Recorded := "FRK_PartRecord"(Core := #Core, Status := #Status, Part := #Part,
                                     RecordName := 'PressDwell', Value := DINT_TO_LREAL(TIME_TO_DINT(#Dwell)), Minimum := 0.0, Maximum := 30000.0,
                                     Target := DINT_TO_LREAL(TIME_TO_DINT(#Dwell)), EngUnit := 'ms');
   END_IF;
   #F_PressDemoRecord := #Core.Exec <> 3;
END_FUNCTION

FUNCTION "FRK_SeqAwait" : Bool   // FC130, SCL
{ S7_Optimized_Access := 'TRUE' }
VERSION : 0.1
// stored: AutoNumber true, IsIECCheckEnabled false, SetENOAutomatically false, UDAEnableTagReadback false
   VAR_INPUT
      Label : String;
      Ok : Bool;
   END_VAR
   VAR_IN_OUT
      Seq : "FRK_SequenceCtx";
   END_VAR
BEGIN

   #FRK_SeqAwait := #Ok;
   IF NOT #Ok AND NOT #Seq.Pending THEN
       #Seq.Pending := TRUE;
       #Seq.Awaiting := #Label;
   END_IF;
END_FUNCTION

